// --- Siemens Structured Format ---
DATA_BLOCK "model_HS16_IW100"
{ S7_Optimized_Access := 'TRUE' }
VERSION : 0.1
NON_RETAIN
   VAR
      W_i : ARRAY[0..15, 0..39] OF REAL;
      W_f : ARRAY[0..15, 0..39] OF REAL;
      W_g : ARRAY[0..15, 0..39] OF REAL;
      W_o : ARRAY[0..15, 0..39] OF REAL;
      R_i : ARRAY[0..15, 0..15] OF REAL;
      R_f : ARRAY[0..15, 0..15] OF REAL;
      R_g : ARRAY[0..15, 0..15] OF REAL;
      R_o : ARRAY[0..15, 0..15] OF REAL;
      B_i : ARRAY[0..15] OF REAL;
      B_f : ARRAY[0..15] OF REAL;
      B_g : ARRAY[0..15] OF REAL;
      B_o : ARRAY[0..15] OF REAL;
      FC_W : ARRAY[0..39, 0..15] OF REAL;
      FC_B : ARRAY[0..39] OF REAL;
   END_VAR
BEGIN

      W_i[0,0] := 0.01364156;
      W_i[0,1] := 0.20536570;
      W_i[0,2] := -0.02245892;
      W_i[0,3] := 0.18291217;
      W_i[0,4] := 0.10548387;
      W_i[0,5] := 0.14748915;
      W_i[0,6] := 0.17824732;
      W_i[0,7] := 0.18831865;
      W_i[0,8] := 0.12917581;
      W_i[0,9] := -0.17035837;
      W_i[0,10] := 0.08922281;
      W_i[0,11] := -0.48598647;
      W_i[0,12] := -0.26934940;
      W_i[0,13] := -0.09021819;
      W_i[0,14] := 0.04866360;
      W_i[0,15] := 0.12027069;
      W_i[0,16] := 0.02211623;
      W_i[0,17] := -0.07331901;
      W_i[0,18] := 0.24969472;
      W_i[0,19] := 0.19951487;
      W_i[0,20] := -0.04635275;
      W_i[0,21] := -0.06017390;
      W_i[0,22] := 0.41972119;
      W_i[0,23] := -0.03179805;
      W_i[0,24] := 0.49648565;
      W_i[0,25] := 0.57860100;
      W_i[0,26] := -0.26113316;
      W_i[0,27] := -0.19300961;
      W_i[0,28] := 0.02716148;
      W_i[0,29] := -0.42831215;
      W_i[0,30] := 0.75518680;
      W_i[0,31] := -0.19160482;
      W_i[0,32] := 0.19652441;
      W_i[0,33] := 0.20859936;
      W_i[0,34] := 0.61514384;
      W_i[0,35] := -0.22654997;
      W_i[0,36] := -0.23919837;
      W_i[0,37] := -0.27295426;
      W_i[0,38] := 0.15717822;
      W_i[0,39] := 0.49166107;
      W_i[1,0] := -0.08388980;
      W_i[1,1] := 0.04137634;
      W_i[1,2] := 0.09732703;
      W_i[1,3] := -0.00114318;
      W_i[1,4] := 0.01266066;
      W_i[1,5] := 0.02146709;
      W_i[1,6] := 0.06203580;
      W_i[1,7] := -0.05510464;
      W_i[1,8] := 0.00995585;
      W_i[1,9] := -0.04009213;
      W_i[1,10] := -0.01534687;
      W_i[1,11] := -0.12621376;
      W_i[1,12] := -0.13568968;
      W_i[1,13] := -0.09674840;
      W_i[1,14] := -0.04467043;
      W_i[1,15] := -0.02089421;
      W_i[1,16] := -0.00725821;
      W_i[1,17] := 0.01724758;
      W_i[1,18] := 0.18129900;
      W_i[1,19] := 0.11187042;
      W_i[1,20] := 0.02454385;
      W_i[1,21] := -0.01102624;
      W_i[1,22] := 0.04567170;
      W_i[1,23] := -0.00008619;
      W_i[1,24] := -0.20038819;
      W_i[1,25] := -0.30851075;
      W_i[1,26] := 0.09543601;
      W_i[1,27] := -0.08277476;
      W_i[1,28] := 0.00373672;
      W_i[1,29] := -0.13582148;
      W_i[1,30] := 0.17890492;
      W_i[1,31] := 0.02590448;
      W_i[1,32] := 0.24079625;
      W_i[1,33] := -0.10525580;
      W_i[1,34] := -0.15286346;
      W_i[1,35] := -0.19629247;
      W_i[1,36] := -0.05740929;
      W_i[1,37] := 0.08565215;
      W_i[1,38] := 0.00725868;
      W_i[1,39] := 0.08298402;
      W_i[2,0] := -0.13536657;
      W_i[2,1] := 0.11532924;
      W_i[2,2] := 0.00179968;
      W_i[2,3] := -0.08932642;
      W_i[2,4] := 0.07508986;
      W_i[2,5] := -0.14212745;
      W_i[2,6] := -0.01394915;
      W_i[2,7] := -0.08767878;
      W_i[2,8] := 0.02846143;
      W_i[2,9] := 0.06891385;
      W_i[2,10] := 0.04481447;
      W_i[2,11] := -0.18693379;
      W_i[2,12] := 0.00844815;
      W_i[2,13] := -0.05949695;
      W_i[2,14] := 0.03289747;
      W_i[2,15] := 0.08402885;
      W_i[2,16] := 0.03656591;
      W_i[2,17] := 0.13008708;
      W_i[2,18] := -0.01728439;
      W_i[2,19] := -0.00760848;
      W_i[2,20] := -0.14490703;
      W_i[2,21] := 0.00184717;
      W_i[2,22] := -0.14345044;
      W_i[2,23] := -0.04114061;
      W_i[2,24] := 0.06368703;
      W_i[2,25] := -0.11341992;
      W_i[2,26] := -0.20044473;
      W_i[2,27] := -0.10808504;
      W_i[2,28] := -0.00091656;
      W_i[2,29] := -0.06285433;
      W_i[2,30] := 0.15420522;
      W_i[2,31] := -0.13147083;
      W_i[2,32] := -0.00983954;
      W_i[2,33] := -0.25118774;
      W_i[2,34] := -0.22324753;
      W_i[2,35] := -0.03245824;
      W_i[2,36] := 0.03434758;
      W_i[2,37] := -0.15230893;
      W_i[2,38] := 0.03214991;
      W_i[2,39] := 0.13666461;
      W_i[3,0] := -0.00015489;
      W_i[3,1] := -0.02602717;
      W_i[3,2] := 0.02940982;
      W_i[3,3] := 0.04201458;
      W_i[3,4] := 0.07303519;
      W_i[3,5] := 0.01782909;
      W_i[3,6] := -0.03795192;
      W_i[3,7] := -0.03116271;
      W_i[3,8] := 0.04315468;
      W_i[3,9] := -0.10355810;
      W_i[3,10] := 0.00910736;
      W_i[3,11] := 0.04493538;
      W_i[3,12] := 0.05511931;
      W_i[3,13] := 0.04794433;
      W_i[3,14] := -0.00690552;
      W_i[3,15] := 0.03096941;
      W_i[3,16] := 0.00754327;
      W_i[3,17] := 0.01626078;
      W_i[3,18] := -0.02028959;
      W_i[3,19] := -0.00735506;
      W_i[3,20] := -0.11980021;
      W_i[3,21] := -0.24100865;
      W_i[3,22] := 0.04234595;
      W_i[3,23] := -0.04032298;
      W_i[3,24] := -0.08977890;
      W_i[3,25] := 0.00863097;
      W_i[3,26] := -0.15812668;
      W_i[3,27] := 0.02937102;
      W_i[3,28] := 0.15920541;
      W_i[3,29] := -0.00798148;
      W_i[3,30] := -0.04935832;
      W_i[3,31] := -0.04004486;
      W_i[3,32] := -0.05156282;
      W_i[3,33] := -0.22839788;
      W_i[3,34] := 0.04730661;
      W_i[3,35] := -0.08628614;
      W_i[3,36] := 0.05156694;
      W_i[3,37] := 0.19403307;
      W_i[3,38] := 0.05496961;
      W_i[3,39] := -0.22899017;
      W_i[4,0] := -0.06762198;
      W_i[4,1] := 0.04105477;
      W_i[4,2] := 0.01412702;
      W_i[4,3] := -0.14503658;
      W_i[4,4] := 0.00052001;
      W_i[4,5] := -0.06361318;
      W_i[4,6] := 0.09927795;
      W_i[4,7] := 0.22318134;
      W_i[4,8] := 0.09787519;
      W_i[4,9] := 0.15435791;
      W_i[4,10] := -0.23381770;
      W_i[4,11] := -0.00151448;
      W_i[4,12] := -0.02443174;
      W_i[4,13] := -0.14362684;
      W_i[4,14] := 0.06250123;
      W_i[4,15] := -0.03108552;
      W_i[4,16] := -0.00760642;
      W_i[4,17] := -0.06110801;
      W_i[4,18] := 0.47297871;
      W_i[4,19] := 0.14145297;
      W_i[4,20] := -0.06666926;
      W_i[4,21] := 0.11880186;
      W_i[4,22] := 0.01305235;
      W_i[4,23] := -0.01088445;
      W_i[4,24] := 0.58226085;
      W_i[4,25] := 0.56463838;
      W_i[4,26] := -0.07272944;
      W_i[4,27] := -0.20381725;
      W_i[4,28] := 0.02941751;
      W_i[4,29] := 0.14696015;
      W_i[4,30] := -0.06698419;
      W_i[4,31] := -0.08342854;
      W_i[4,32] := 0.09379109;
      W_i[4,33] := 0.14583473;
      W_i[4,34] := -0.02093923;
      W_i[4,35] := -0.13240194;
      W_i[4,36] := -0.03764428;
      W_i[4,37] := -0.08758924;
      W_i[4,38] := -0.06055138;
      W_i[4,39] := 0.54854435;
      W_i[5,0] := -0.26418173;
      W_i[5,1] := 0.00919414;
      W_i[5,2] := 0.28921035;
      W_i[5,3] := 0.19848731;
      W_i[5,4] := 0.04857918;
      W_i[5,5] := -0.07696015;
      W_i[5,6] := -0.18773772;
      W_i[5,7] := -0.06413802;
      W_i[5,8] := -0.19999725;
      W_i[5,9] := 0.00090761;
      W_i[5,10] := 0.06217722;
      W_i[5,11] := 0.10535000;
      W_i[5,12] := -0.20478797;
      W_i[5,13] := 0.00378444;
      W_i[5,14] := -0.08047202;
      W_i[5,15] := 0.10188833;
      W_i[5,16] := -0.10373244;
      W_i[5,17] := 0.02060685;
      W_i[5,18] := 0.26179335;
      W_i[5,19] := -0.16465248;
      W_i[5,20] := -0.21371244;
      W_i[5,21] := 0.18068251;
      W_i[5,22] := -0.14789225;
      W_i[5,23] := -0.00876896;
      W_i[5,24] := 0.22973008;
      W_i[5,25] := 0.59550780;
      W_i[5,26] := 0.14612897;
      W_i[5,27] := -0.08599184;
      W_i[5,28] := -0.22050266;
      W_i[5,29] := -0.17621692;
      W_i[5,30] := -0.21464045;
      W_i[5,31] := -0.01781221;
      W_i[5,32] := -0.06129935;
      W_i[5,33] := 0.05988304;
      W_i[5,34] := 0.25511330;
      W_i[5,35] := -0.14653285;
      W_i[5,36] := -0.15237394;
      W_i[5,37] := -0.39873159;
      W_i[5,38] := 0.06444512;
      W_i[5,39] := -0.46595329;
      W_i[6,0] := -0.09987911;
      W_i[6,1] := -0.35666752;
      W_i[6,2] := -0.14997965;
      W_i[6,3] := -0.16122143;
      W_i[6,4] := -0.03222676;
      W_i[6,5] := -0.06696601;
      W_i[6,6] := -0.18053886;
      W_i[6,7] := -0.38125506;
      W_i[6,8] := 0.15195245;
      W_i[6,9] := -0.12253319;
      W_i[6,10] := -0.06935552;
      W_i[6,11] := -0.25237226;
      W_i[6,12] := -0.00955063;
      W_i[6,13] := -0.13364333;
      W_i[6,14] := 0.12441263;
      W_i[6,15] := -0.06698428;
      W_i[6,16] := 0.02953966;
      W_i[6,17] := -0.12817322;
      W_i[6,18] := 0.50510013;
      W_i[6,19] := -0.07000107;
      W_i[6,20] := 0.10518134;
      W_i[6,21] := -0.12933129;
      W_i[6,22] := 0.08060265;
      W_i[6,23] := 0.16216518;
      W_i[6,24] := 0.56379879;
      W_i[6,25] := 0.51589292;
      W_i[6,26] := -0.06017810;
      W_i[6,27] := 0.13627745;
      W_i[6,28] := 0.07406422;
      W_i[6,29] := -0.04566135;
      W_i[6,30] := 0.11365223;
      W_i[6,31] := -0.19966318;
      W_i[6,32] := 0.05134548;
      W_i[6,33] := -0.06383436;
      W_i[6,34] := 0.18601419;
      W_i[6,35] := -0.00495438;
      W_i[6,36] := -0.01991113;
      W_i[6,37] := 0.13569827;
      W_i[6,38] := 0.10721204;
      W_i[6,39] := -0.19543035;
      W_i[7,0] := 0.11805627;
      W_i[7,1] := 0.06404518;
      W_i[7,2] := 0.26091906;
      W_i[7,3] := -0.13242221;
      W_i[7,4] := 0.04345745;
      W_i[7,5] := 0.06463753;
      W_i[7,6] := 0.14174174;
      W_i[7,7] := 0.17861204;
      W_i[7,8] := 0.14897110;
      W_i[7,9] := -0.10119636;
      W_i[7,10] := -0.21339175;
      W_i[7,11] := -0.29427007;
      W_i[7,12] := -0.12524955;
      W_i[7,13] := -0.22747980;
      W_i[7,14] := -0.08303443;
      W_i[7,15] := 0.15086012;
      W_i[7,16] := -0.02865510;
      W_i[7,17] := 0.14286377;
      W_i[7,18] := 0.06569705;
      W_i[7,19] := 0.17024888;
      W_i[7,20] := 0.16341139;
      W_i[7,21] := -0.08116058;
      W_i[7,22] := 0.28119785;
      W_i[7,23] := -0.24578308;
      W_i[7,24] := 0.46118793;
      W_i[7,25] := 0.87448853;
      W_i[7,26] := -0.21451366;
      W_i[7,27] := -0.03196089;
      W_i[7,28] := 0.11030190;
      W_i[7,29] := 0.08675592;
      W_i[7,30] := 0.63182199;
      W_i[7,31] := 0.09978309;
      W_i[7,32] := -0.11112560;
      W_i[7,33] := 0.14244974;
      W_i[7,34] := 0.87706214;
      W_i[7,35] := 0.04549777;
      W_i[7,36] := 0.01875403;
      W_i[7,37] := 0.19351047;
      W_i[7,38] := 0.04132079;
      W_i[7,39] := 0.30163178;
      W_i[8,0] := 0.00448507;
      W_i[8,1] := 0.00593045;
      W_i[8,2] := 0.05385492;
      W_i[8,3] := 0.23692533;
      W_i[8,4] := 0.13600577;
      W_i[8,5] := -0.13479330;
      W_i[8,6] := 0.05155064;
      W_i[8,7] := -0.18396251;
      W_i[8,8] := -0.04175631;
      W_i[8,9] := 0.02508196;
      W_i[8,10] := 0.08028799;
      W_i[8,11] := -0.09709663;
      W_i[8,12] := -0.24632221;
      W_i[8,13] := -0.09933189;
      W_i[8,14] := -0.13090380;
      W_i[8,15] := 0.08873132;
      W_i[8,16] := -0.15212885;
      W_i[8,17] := 0.09358153;
      W_i[8,18] := -0.04925272;
      W_i[8,19] := -0.20840898;
      W_i[8,20] := -0.08381097;
      W_i[8,21] := 0.06258945;
      W_i[8,22] := -0.07553499;
      W_i[8,23] := -0.05963936;
      W_i[8,24] := 0.35542277;
      W_i[8,25] := 0.42086950;
      W_i[8,26] := 0.08319889;
      W_i[8,27] := -0.18197235;
      W_i[8,28] := 0.06505518;
      W_i[8,29] := 0.07391432;
      W_i[8,30] := 0.12715283;
      W_i[8,31] := -0.13722460;
      W_i[8,32] := 0.24457708;
      W_i[8,33] := 0.17096752;
      W_i[8,34] := -0.13092747;
      W_i[8,35] := 0.11238978;
      W_i[8,36] := -0.01007767;
      W_i[8,37] := 0.04878357;
      W_i[8,38] := -0.09178042;
      W_i[8,39] := 0.70590818;
      W_i[9,0] := 0.13898331;
      W_i[9,1] := 0.21558045;
      W_i[9,2] := -0.01587300;
      W_i[9,3] := -0.02008759;
      W_i[9,4] := 0.14031912;
      W_i[9,5] := 0.14432517;
      W_i[9,6] := 0.22022982;
      W_i[9,7] := 0.11039817;
      W_i[9,8] := -0.01799948;
      W_i[9,9] := 0.01688460;
      W_i[9,10] := 0.08939565;
      W_i[9,11] := 0.15729012;
      W_i[9,12] := -0.16055229;
      W_i[9,13] := 0.07329134;
      W_i[9,14] := 0.03671210;
      W_i[9,15] := 0.07092312;
      W_i[9,16] := -0.01012265;
      W_i[9,17] := 0.03808835;
      W_i[9,18] := -0.00362916;
      W_i[9,19] := -0.00791038;
      W_i[9,20] := 0.13901256;
      W_i[9,21] := -0.05212758;
      W_i[9,22] := -0.13945961;
      W_i[9,23] := 0.01820100;
      W_i[9,24] := -0.28223145;
      W_i[9,25] := -0.05683075;
      W_i[9,26] := -0.06647032;
      W_i[9,27] := 0.11427623;
      W_i[9,28] := -0.05756322;
      W_i[9,29] := 0.25496486;
      W_i[9,30] := -0.41661564;
      W_i[9,31] := 0.03821095;
      W_i[9,32] := -0.24074574;
      W_i[9,33] := -0.01633074;
      W_i[9,34] := -0.30772033;
      W_i[9,35] := -0.30636224;
      W_i[9,36] := -0.00646075;
      W_i[9,37] := -0.10956979;
      W_i[9,38] := 0.04284515;
      W_i[9,39] := 0.06388737;
      W_i[10,0] := 0.15491682;
      W_i[10,1] := 0.06016659;
      W_i[10,2] := 0.08790326;
      W_i[10,3] := 0.04701571;
      W_i[10,4] := -0.21938066;
      W_i[10,5] := -0.00418864;
      W_i[10,6] := -0.14329411;
      W_i[10,7] := -0.13763005;
      W_i[10,8] := -0.07890343;
      W_i[10,9] := 0.10256134;
      W_i[10,10] := -0.02710062;
      W_i[10,11] := -0.20991582;
      W_i[10,12] := 0.43801337;
      W_i[10,13] := 0.07667056;
      W_i[10,14] := -0.05265489;
      W_i[10,15] := 0.09571737;
      W_i[10,16] := -0.14256968;
      W_i[10,17] := 0.00645238;
      W_i[10,18] := 0.08263779;
      W_i[10,19] := -0.13588426;
      W_i[10,20] := 0.17050405;
      W_i[10,21] := 0.34270245;
      W_i[10,22] := 0.12177468;
      W_i[10,23] := 0.03954393;
      W_i[10,24] := 0.78272396;
      W_i[10,25] := 0.62249583;
      W_i[10,26] := -0.04197677;
      W_i[10,27] := -0.01324140;
      W_i[10,28] := -0.11742962;
      W_i[10,29] := 0.03315270;
      W_i[10,30] := 0.43726227;
      W_i[10,31] := -0.01188345;
      W_i[10,32] := 0.02015782;
      W_i[10,33] := 0.26254645;
      W_i[10,34] := 0.31372723;
      W_i[10,35] := 0.13515088;
      W_i[10,36] := -0.13856903;
      W_i[10,37] := -0.07906500;
      W_i[10,38] := 0.04151168;
      W_i[10,39] := 0.58438212;
      W_i[11,0] := -0.03692184;
      W_i[11,1] := 0.08602915;
      W_i[11,2] := 0.04734402;
      W_i[11,3] := 0.15488507;
      W_i[11,4] := 0.02953814;
      W_i[11,5] := -0.03516553;
      W_i[11,6] := -0.03630468;
      W_i[11,7] := 0.22055247;
      W_i[11,8] := 0.05422686;
      W_i[11,9] := -0.19223477;
      W_i[11,10] := 0.15922990;
      W_i[11,11] := -0.50660896;
      W_i[11,12] := 0.21863456;
      W_i[11,13] := 0.06115106;
      W_i[11,14] := 0.05269584;
      W_i[11,15] := 0.01791226;
      W_i[11,16] := -0.08076685;
      W_i[11,17] := -0.00192191;
      W_i[11,18] := 0.20004040;
      W_i[11,19] := -0.02625836;
      W_i[11,20] := 0.02325124;
      W_i[11,21] := 0.02411360;
      W_i[11,22] := -0.03470324;
      W_i[11,23] := 0.02441446;
      W_i[11,24] := 0.01363192;
      W_i[11,25] := -0.20787865;
      W_i[11,26] := -0.09482310;
      W_i[11,27] := 0.05317536;
      W_i[11,28] := 0.01368785;
      W_i[11,29] := 0.24679546;
      W_i[11,30] := 0.09310606;
      W_i[11,31] := 0.02022941;
      W_i[11,32] := 0.25092661;
      W_i[11,33] := -0.02307699;
      W_i[11,34] := -0.18370298;
      W_i[11,35] := 0.24884717;
      W_i[11,36] := -0.08544295;
      W_i[11,37] := -0.04159483;
      W_i[11,38] := 0.12627473;
      W_i[11,39] := 0.57147032;
      W_i[12,0] := 0.26667652;
      W_i[12,1] := 0.18141651;
      W_i[12,2] := -0.04977122;
      W_i[12,3] := 0.09079568;
      W_i[12,4] := 0.22469823;
      W_i[12,5] := -0.13473749;
      W_i[12,6] := 0.22730011;
      W_i[12,7] := -0.10648373;
      W_i[12,8] := 0.00375756;
      W_i[12,9] := 0.14409521;
      W_i[12,10] := -0.04439257;
      W_i[12,11] := 0.01341529;
      W_i[12,12] := 0.05264389;
      W_i[12,13] := 0.14714998;
      W_i[12,14] := 0.02812583;
      W_i[12,15] := 0.09371702;
      W_i[12,16] := -0.01640923;
      W_i[12,17] := -0.00820156;
      W_i[12,18] := -0.02099935;
      W_i[12,19] := 0.03455377;
      W_i[12,20] := -0.00376845;
      W_i[12,21] := 0.01287318;
      W_i[12,22] := 0.27967688;
      W_i[12,23] := 0.32648781;
      W_i[12,24] := -0.04639676;
      W_i[12,25] := -0.12604533;
      W_i[12,26] := -0.05218698;
      W_i[12,27] := 0.19303280;
      W_i[12,28] := -0.02861599;
      W_i[12,29] := 0.07526918;
      W_i[12,30] := 0.27195212;
      W_i[12,31] := -0.24740550;
      W_i[12,32] := 0.12962508;
      W_i[12,33] := -0.02061021;
      W_i[12,34] := -0.38526946;
      W_i[12,35] := -0.44955108;
      W_i[12,36] := 0.17704585;
      W_i[12,37] := -0.58847874;
      W_i[12,38] := 0.02093910;
      W_i[12,39] := -0.07715891;
      W_i[13,0] := 0.02638375;
      W_i[13,1] := 0.04267908;
      W_i[13,2] := -0.04100905;
      W_i[13,3] := 0.02433234;
      W_i[13,4] := 0.19633174;
      W_i[13,5] := 0.09253235;
      W_i[13,6] := 0.18767522;
      W_i[13,7] := -0.09313158;
      W_i[13,8] := 0.06435700;
      W_i[13,9] := -0.02719559;
      W_i[13,10] := 0.11561871;
      W_i[13,11] := -0.12066963;
      W_i[13,12] := -0.27772844;
      W_i[13,13] := -0.00763909;
      W_i[13,14] := 0.07759997;
      W_i[13,15] := 0.01202866;
      W_i[13,16] := 0.07374192;
      W_i[13,17] := 0.03084671;
      W_i[13,18] := -0.03566260;
      W_i[13,19] := 0.21000803;
      W_i[13,20] := -0.08411094;
      W_i[13,21] := -0.21406713;
      W_i[13,22] := 0.03648549;
      W_i[13,23] := -0.03847607;
      W_i[13,24] := 0.70946354;
      W_i[13,25] := 0.49792659;
      W_i[13,26] := -0.08645725;
      W_i[13,27] := 0.15172665;
      W_i[13,28] := -0.01545484;
      W_i[13,29] := 0.07564367;
      W_i[13,30] := 0.04488704;
      W_i[13,31] := -0.05433368;
      W_i[13,32] := -0.12254967;
      W_i[13,33] := 0.05323875;
      W_i[13,34] := 0.28031611;
      W_i[13,35] := -0.31686431;
      W_i[13,36] := 0.08479394;
      W_i[13,37] := -0.18495709;
      W_i[13,38] := 0.10758790;
      W_i[13,39] := 0.68741995;
      W_i[14,0] := -0.17416088;
      W_i[14,1] := 0.01005446;
      W_i[14,2] := -0.26855752;
      W_i[14,3] := -0.62796623;
      W_i[14,4] := 0.06820592;
      W_i[14,5] := -0.16153112;
      W_i[14,6] := 0.04283209;
      W_i[14,7] := -0.29056939;
      W_i[14,8] := -0.67249602;
      W_i[14,9] := -0.34167016;
      W_i[14,10] := 0.09426845;
      W_i[14,11] := -0.10104106;
      W_i[14,12] := 0.10796092;
      W_i[14,13] := -0.18351264;
      W_i[14,14] := 0.00065603;
      W_i[14,15] := -0.06139126;
      W_i[14,16] := -0.11547680;
      W_i[14,17] := 0.04488576;
      W_i[14,18] := -0.15664500;
      W_i[14,19] := 0.00779267;
      W_i[14,20] := -0.01367023;
      W_i[14,21] := -0.02746255;
      W_i[14,22] := -0.06486769;
      W_i[14,23] := 0.17152609;
      W_i[14,24] := -0.10990940;
      W_i[14,25] := -0.08006914;
      W_i[14,26] := -0.25285053;
      W_i[14,27] := 0.06160279;
      W_i[14,28] := 0.17719766;
      W_i[14,29] := 0.14922956;
      W_i[14,30] := 0.00092594;
      W_i[14,31] := -0.11380912;
      W_i[14,32] := -0.09275766;
      W_i[14,33] := -0.05691696;
      W_i[14,34] := -0.20431529;
      W_i[14,35] := -0.06423868;
      W_i[14,36] := -0.08797362;
      W_i[14,37] := -0.07569788;
      W_i[14,38] := 0.23112053;
      W_i[14,39] := 0.00680392;
      W_i[15,0] := 0.02184013;
      W_i[15,1] := 0.18801539;
      W_i[15,2] := 0.06529985;
      W_i[15,3] := -0.13560045;
      W_i[15,4] := 0.14931200;
      W_i[15,5] := -0.07038850;
      W_i[15,6] := -0.03877895;
      W_i[15,7] := 0.08169580;
      W_i[15,8] := 0.04022081;
      W_i[15,9] := 0.16485462;
      W_i[15,10] := 0.02359114;
      W_i[15,11] := -0.06464480;
      W_i[15,12] := -0.13054129;
      W_i[15,13] := 0.14513132;
      W_i[15,14] := -0.00291753;
      W_i[15,15] := 0.00511506;
      W_i[15,16] := 0.04386861;
      W_i[15,17] := -0.14875175;
      W_i[15,18] := -0.02457544;
      W_i[15,19] := 0.07704978;
      W_i[15,20] := -0.04825005;
      W_i[15,21] := 0.03190987;
      W_i[15,22] := -0.09410153;
      W_i[15,23] := -0.16679235;
      W_i[15,24] := -0.46764547;
      W_i[15,25] := -0.44318548;
      W_i[15,26] := -0.05940514;
      W_i[15,27] := 0.05163483;
      W_i[15,28] := -0.03008339;
      W_i[15,29] := 0.21256405;
      W_i[15,30] := -0.05510921;
      W_i[15,31] := -0.09820909;
      W_i[15,32] := 0.21482152;
      W_i[15,33] := 0.30279014;
      W_i[15,34] := -0.06246981;
      W_i[15,35] := 0.01027228;
      W_i[15,36] := -0.09376621;
      W_i[15,37] := -0.02936010;
      W_i[15,38] := -0.47935137;
      W_i[15,39] := 0.05519279;
      W_f[0,0] := 0.05364275;
      W_f[0,1] := 0.09687193;
      W_f[0,2] := -0.03420604;
      W_f[0,3] := 0.09112332;
      W_f[0,4] := 0.01952212;
      W_f[0,5] := -0.00599490;
      W_f[0,6] := -0.02583287;
      W_f[0,7] := 0.01641575;
      W_f[0,8] := 0.00249371;
      W_f[0,9] := -0.03082566;
      W_f[0,10] := 0.03822958;
      W_f[0,11] := -0.20525688;
      W_f[0,12] := 0.15610816;
      W_f[0,13] := 0.01319965;
      W_f[0,14] := -0.00955972;
      W_f[0,15] := -0.01736578;
      W_f[0,16] := -0.01232213;
      W_f[0,17] := -0.07847971;
      W_f[0,18] := 0.03267125;
      W_f[0,19] := 0.02281226;
      W_f[0,20] := -0.00946235;
      W_f[0,21] := -0.04914912;
      W_f[0,22] := -0.05509606;
      W_f[0,23] := -0.04103199;
      W_f[0,24] := 0.49705139;
      W_f[0,25] := 0.41528228;
      W_f[0,26] := -0.10808732;
      W_f[0,27] := -0.04818393;
      W_f[0,28] := 0.06444012;
      W_f[0,29] := -0.15780614;
      W_f[0,30] := 0.10075731;
      W_f[0,31] := -0.03347747;
      W_f[0,32] := 0.13920051;
      W_f[0,33] := -0.07730422;
      W_f[0,34] := 0.22286199;
      W_f[0,35] := 0.09730371;
      W_f[0,36] := 0.01644731;
      W_f[0,37] := -0.14617991;
      W_f[0,38] := -0.03747354;
      W_f[0,39] := 0.08508820;
      W_f[1,0] := -0.03535822;
      W_f[1,1] := -0.47124356;
      W_f[1,2] := -0.14644240;
      W_f[1,3] := 0.07842869;
      W_f[1,4] := -0.00283514;
      W_f[1,5] := 0.13242532;
      W_f[1,6] := -0.17787769;
      W_f[1,7] := 0.03437876;
      W_f[1,8] := -0.30326170;
      W_f[1,9] := 0.03390699;
      W_f[1,10] := 0.04835700;
      W_f[1,11] := 0.39755464;
      W_f[1,12] := 0.22270909;
      W_f[1,13] := 0.21808504;
      W_f[1,14] := -0.11776564;
      W_f[1,15] := 0.10067453;
      W_f[1,16] := -0.36373556;
      W_f[1,17] := 0.18559641;
      W_f[1,18] := 0.40969753;
      W_f[1,19] := 0.12707092;
      W_f[1,20] := 0.29767519;
      W_f[1,21] := -0.16713570;
      W_f[1,22] := -0.17408817;
      W_f[1,23] := 0.12793775;
      W_f[1,24] := -0.53485709;
      W_f[1,25] := -0.56272870;
      W_f[1,26] := 0.05998780;
      W_f[1,27] := 0.01051460;
      W_f[1,28] := -0.12135706;
      W_f[1,29] := 0.13744721;
      W_f[1,30] := -0.09007506;
      W_f[1,31] := -0.00778998;
      W_f[1,32] := 0.11112776;
      W_f[1,33] := -0.16928056;
      W_f[1,34] := 0.31107175;
      W_f[1,35] := 0.19411123;
      W_f[1,36] := -0.06959353;
      W_f[1,37] := -0.25251710;
      W_f[1,38] := 0.34865397;
      W_f[1,39] := 0.05812330;
      W_f[2,0] := -0.03221922;
      W_f[2,1] := 0.12347551;
      W_f[2,2] := -0.06227477;
      W_f[2,3] := 0.20185524;
      W_f[2,4] := 0.00543583;
      W_f[2,5] := 0.03781491;
      W_f[2,6] := -0.00314693;
      W_f[2,7] := 0.04292703;
      W_f[2,8] := -0.00575330;
      W_f[2,9] := -0.08594991;
      W_f[2,10] := -0.01364730;
      W_f[2,11] := -0.17743753;
      W_f[2,12] := -0.00461064;
      W_f[2,13] := -0.05826429;
      W_f[2,14] := 0.06936967;
      W_f[2,15] := 0.02028695;
      W_f[2,16] := 0.00601915;
      W_f[2,17] := 0.02327365;
      W_f[2,18] := -0.03857812;
      W_f[2,19] := -0.08794222;
      W_f[2,20] := 0.01833609;
      W_f[2,21] := 0.03344638;
      W_f[2,22] := -0.09674103;
      W_f[2,23] := 0.03481310;
      W_f[2,24] := -0.20710675;
      W_f[2,25] := -0.12916997;
      W_f[2,26] := 0.00745270;
      W_f[2,27] := -0.01033618;
      W_f[2,28] := 0.07703895;
      W_f[2,29] := 0.08949607;
      W_f[2,30] := -0.07744866;
      W_f[2,31] := -0.00363669;
      W_f[2,32] := -0.10897757;
      W_f[2,33] := 0.05933027;
      W_f[2,34] := 0.12423457;
      W_f[2,35] := -0.08927383;
      W_f[2,36] := -0.00645528;
      W_f[2,37] := 0.19684052;
      W_f[2,38] := -0.12688994;
      W_f[2,39] := 0.15507455;
      W_f[3,0] := -0.15219240;
      W_f[3,1] := -0.09112048;
      W_f[3,2] := -0.13655797;
      W_f[3,3] := 0.09398650;
      W_f[3,4] := -0.38095236;
      W_f[3,5] := 0.07147726;
      W_f[3,6] := 0.27381626;
      W_f[3,7] := -0.03780884;
      W_f[3,8] := -0.09247751;
      W_f[3,9] := 0.32965410;
      W_f[3,10] := -0.21033977;
      W_f[3,11] := -0.01770502;
      W_f[3,12] := -0.16563010;
      W_f[3,13] := -0.09659225;
      W_f[3,14] := -0.14708968;
      W_f[3,15] := -0.04307340;
      W_f[3,16] := -0.04020571;
      W_f[3,17] := -0.15388337;
      W_f[3,18] := 0.04561477;
      W_f[3,19] := -0.03800451;
      W_f[3,20] := -0.11640513;
      W_f[3,21] := 0.10628393;
      W_f[3,22] := 0.13051899;
      W_f[3,23] := 0.15934397;
      W_f[3,24] := -0.49496132;
      W_f[3,25] := -0.46555015;
      W_f[3,26] := 0.07467606;
      W_f[3,27] := 0.05813665;
      W_f[3,28] := -0.45595208;
      W_f[3,29] := 0.13731937;
      W_f[3,30] := -0.04639205;
      W_f[3,31] := 0.20856442;
      W_f[3,32] := 0.23197061;
      W_f[3,33] := -0.09503688;
      W_f[3,34] := 0.22798222;
      W_f[3,35] := -0.10183924;
      W_f[3,36] := 0.24291022;
      W_f[3,37] := 0.09243517;
      W_f[3,38] := -0.01472234;
      W_f[3,39] := 0.84467447;
      W_f[4,0] := 0.02846950;
      W_f[4,1] := 0.06578626;
      W_f[4,2] := 0.00272045;
      W_f[4,3] := 0.02383544;
      W_f[4,4] := -0.04941020;
      W_f[4,5] := 0.03107557;
      W_f[4,6] := 0.04498140;
      W_f[4,7] := 0.00715393;
      W_f[4,8] := -0.00156786;
      W_f[4,9] := 0.01842991;
      W_f[4,10] := -0.02190995;
      W_f[4,11] := 0.00170467;
      W_f[4,12] := -0.11754189;
      W_f[4,13] := -0.00572082;
      W_f[4,14] := -0.02148229;
      W_f[4,15] := -0.02594547;
      W_f[4,16] := -0.06025682;
      W_f[4,17] := -0.08476730;
      W_f[4,18] := 0.07604560;
      W_f[4,19] := 0.05858169;
      W_f[4,20] := 0.05974808;
      W_f[4,21] := 0.24128842;
      W_f[4,22] := 0.16804713;
      W_f[4,23] := -0.03820573;
      W_f[4,24] := 0.48765618;
      W_f[4,25] := 0.57080442;
      W_f[4,26] := -0.00810769;
      W_f[4,27] := -0.18718927;
      W_f[4,28] := 0.06110260;
      W_f[4,29] := -0.09344726;
      W_f[4,30] := 0.46467450;
      W_f[4,31] := 0.05612971;
      W_f[4,32] := 0.03677486;
      W_f[4,33] := 0.11877728;
      W_f[4,34] := 0.03321171;
      W_f[4,35] := 0.29353175;
      W_f[4,36] := 0.05504971;
      W_f[4,37] := 0.10279266;
      W_f[4,38] := -0.00283241;
      W_f[4,39] := 0.06622307;
      W_f[5,0] := 0.11376505;
      W_f[5,1] := 0.04806940;
      W_f[5,2] := -0.10279931;
      W_f[5,3] := -0.16593064;
      W_f[5,4] := 0.00000844;
      W_f[5,5] := 0.02789909;
      W_f[5,6] := 0.04521109;
      W_f[5,7] := 0.02275284;
      W_f[5,8] := -0.02738458;
      W_f[5,9] := 0.06878603;
      W_f[5,10] := -0.01160701;
      W_f[5,11] := -0.05195494;
      W_f[5,12] := -0.10548418;
      W_f[5,13] := 0.01500680;
      W_f[5,14] := 0.08265527;
      W_f[5,15] := 0.00386744;
      W_f[5,16] := 0.05198263;
      W_f[5,17] := 0.02937749;
      W_f[5,18] := 0.06512810;
      W_f[5,19] := 0.03703250;
      W_f[5,20] := 0.06421617;
      W_f[5,21] := -0.01455062;
      W_f[5,22] := 0.19789651;
      W_f[5,23] := -0.03008014;
      W_f[5,24] := 0.34697571;
      W_f[5,25] := 0.65106732;
      W_f[5,26] := -0.00135605;
      W_f[5,27] := 0.05647351;
      W_f[5,28] := 0.09934321;
      W_f[5,29] := -0.13159826;
      W_f[5,30] := 0.01969404;
      W_f[5,31] := 0.03655320;
      W_f[5,32] := -0.05406484;
      W_f[5,33] := -0.11042146;
      W_f[5,34] := 0.09479982;
      W_f[5,35] := 0.04922118;
      W_f[5,36] := 0.04102103;
      W_f[5,37] := 0.20328595;
      W_f[5,38] := 0.09994788;
      W_f[5,39] := 0.16133195;
      W_f[6,0] := -0.03485869;
      W_f[6,1] := -0.00908120;
      W_f[6,2] := -0.03699812;
      W_f[6,3] := -0.03682025;
      W_f[6,4] := 0.09187597;
      W_f[6,5] := 0.05246547;
      W_f[6,6] := 0.12492345;
      W_f[6,7] := -0.00999346;
      W_f[6,8] := -0.08344354;
      W_f[6,9] := 0.07932125;
      W_f[6,10] := 0.03438351;
      W_f[6,11] := -0.06988891;
      W_f[6,12] := 0.03135443;
      W_f[6,13] := 0.00137540;
      W_f[6,14] := 0.03249843;
      W_f[6,15] := -0.01266906;
      W_f[6,16] := -0.00345383;
      W_f[6,17] := -0.07384243;
      W_f[6,18] := -0.04767740;
      W_f[6,19] := 0.00589593;
      W_f[6,20] := 0.04428503;
      W_f[6,21] := 0.05965255;
      W_f[6,22] := 0.13275859;
      W_f[6,23] := -0.07216866;
      W_f[6,24] := 0.32743850;
      W_f[6,25] := 0.41480702;
      W_f[6,26] := 0.00211261;
      W_f[6,27] := -0.02340442;
      W_f[6,28] := -0.04405304;
      W_f[6,29] := 0.02433619;
      W_f[6,30] := -0.18997696;
      W_f[6,31] := 0.13028599;
      W_f[6,32] := 0.16898793;
      W_f[6,33] := 0.09330611;
      W_f[6,34] := 0.04484965;
      W_f[6,35] := -0.08660950;
      W_f[6,36] := -0.02266579;
      W_f[6,37] := 0.11412326;
      W_f[6,38] := 0.07686570;
      W_f[6,39] := -0.11869525;
      W_f[7,0] := -0.00221147;
      W_f[7,1] := 0.10511280;
      W_f[7,2] := -0.07019065;
      W_f[7,3] := -0.01243510;
      W_f[7,4] := 0.02943816;
      W_f[7,5] := 0.06614972;
      W_f[7,6] := 0.04611924;
      W_f[7,7] := 0.02763495;
      W_f[7,8] := -0.01057697;
      W_f[7,9] := -0.02540869;
      W_f[7,10] := -0.00237630;
      W_f[7,11] := -0.14796597;
      W_f[7,12] := 0.04395492;
      W_f[7,13] := 0.07364006;
      W_f[7,14] := -0.03409544;
      W_f[7,15] := -0.07690118;
      W_f[7,16] := 0.00728678;
      W_f[7,17] := 0.07319640;
      W_f[7,18] := 0.06380690;
      W_f[7,19] := 0.00555583;
      W_f[7,20] := -0.01266172;
      W_f[7,21] := 0.05246431;
      W_f[7,22] := 0.13432735;
      W_f[7,23] := 0.00786275;
      W_f[7,24] := 0.36037040;
      W_f[7,25] := 0.63975710;
      W_f[7,26] := -0.14318357;
      W_f[7,27] := 0.02217500;
      W_f[7,28] := 0.03329759;
      W_f[7,29] := 0.02024308;
      W_f[7,30] := 0.06194379;
      W_f[7,31] := -0.03574094;
      W_f[7,32] := 0.27383688;
      W_f[7,33] := 0.09022309;
      W_f[7,34] := 0.72298384;
      W_f[7,35] := -0.13958853;
      W_f[7,36] := -0.05832926;
      W_f[7,37] := 0.05806842;
      W_f[7,38] := 0.01794156;
      W_f[7,39] := 0.00930902;
      W_f[8,0] := -0.00069194;
      W_f[8,1] := 0.09570718;
      W_f[8,2] := -0.13032150;
      W_f[8,3] := -0.00169487;
      W_f[8,4] := 0.05343744;
      W_f[8,5] := 0.05416366;
      W_f[8,6] := 0.00489102;
      W_f[8,7] := 0.04302023;
      W_f[8,8] := 0.02923981;
      W_f[8,9] := -0.03308041;
      W_f[8,10] := 0.02764279;
      W_f[8,11] := -0.08082840;
      W_f[8,12] := -0.04773318;
      W_f[8,13] := -0.02026195;
      W_f[8,14] := -0.02248771;
      W_f[8,15] := -0.14968230;
      W_f[8,16] := 0.10387620;
      W_f[8,17] := 0.02660801;
      W_f[8,18] := 0.02133987;
      W_f[8,19] := 0.06662087;
      W_f[8,20] := 0.02782230;
      W_f[8,21] := 0.01667393;
      W_f[8,22] := 0.29885378;
      W_f[8,23] := -0.04644651;
      W_f[8,24] := 0.36805248;
      W_f[8,25] := 0.58228642;
      W_f[8,26] := -0.01743001;
      W_f[8,27] := -0.01691605;
      W_f[8,28] := 0.01118935;
      W_f[8,29] := -0.00426544;
      W_f[8,30] := 0.17033555;
      W_f[8,31] := -0.03053380;
      W_f[8,32] := 0.12107975;
      W_f[8,33] := -0.06191333;
      W_f[8,34] := 0.74060959;
      W_f[8,35] := -0.07475549;
      W_f[8,36] := -0.02023359;
      W_f[8,37] := 0.02331678;
      W_f[8,38] := -0.03007067;
      W_f[8,39] := -0.05748938;
      W_f[9,0] := -0.10508082;
      W_f[9,1] := -0.04133019;
      W_f[9,2] := -0.06146885;
      W_f[9,3] := 0.03741426;
      W_f[9,4] := -0.08707085;
      W_f[9,5] := -0.06223321;
      W_f[9,6] := -0.18814664;
      W_f[9,7] := -0.11111913;
      W_f[9,8] := -0.13546698;
      W_f[9,9] := -0.00564482;
      W_f[9,10] := -0.01552745;
      W_f[9,11] := -0.17684816;
      W_f[9,12] := 0.03565479;
      W_f[9,13] := -0.08725277;
      W_f[9,14] := -0.00522599;
      W_f[9,15] := -0.10947887;
      W_f[9,16] := 0.01476094;
      W_f[9,17] := -0.05979283;
      W_f[9,18] := -0.00063397;
      W_f[9,19] := 0.06166672;
      W_f[9,20] := -0.10422222;
      W_f[9,21] := 0.00166027;
      W_f[9,22] := -0.27992189;
      W_f[9,23] := -0.03734995;
      W_f[9,24] := 0.12155679;
      W_f[9,25] := -0.06815521;
      W_f[9,26] := -0.01121978;
      W_f[9,27] := -0.01608659;
      W_f[9,28] := 0.04067907;
      W_f[9,29] := -0.06756267;
      W_f[9,30] := 0.05508788;
      W_f[9,31] := -0.09057643;
      W_f[9,32] := -0.07261790;
      W_f[9,33] := -0.13291492;
      W_f[9,34] := -0.02277668;
      W_f[9,35] := 0.19900511;
      W_f[9,36] := -0.00467835;
      W_f[9,37] := -0.18864036;
      W_f[9,38] := 0.01334353;
      W_f[9,39] := -0.01253361;
      W_f[10,0] := -0.00524171;
      W_f[10,1] := 0.10620133;
      W_f[10,2] := -0.06919775;
      W_f[10,3] := -0.00134773;
      W_f[10,4] := -0.01228707;
      W_f[10,5] := 0.01736076;
      W_f[10,6] := 0.03687445;
      W_f[10,7] := 0.02915340;
      W_f[10,8] := 0.06300525;
      W_f[10,9] := -0.06548626;
      W_f[10,10] := 0.05580841;
      W_f[10,11] := -0.10701931;
      W_f[10,12] := -0.02223501;
      W_f[10,13] := 0.00853262;
      W_f[10,14] := 0.03023283;
      W_f[10,15] := -0.06348655;
      W_f[10,16] := 0.04187576;
      W_f[10,17] := 0.00731900;
      W_f[10,18] := 0.08542238;
      W_f[10,19] := 0.00890474;
      W_f[10,20] := 0.07895420;
      W_f[10,21] := 0.07658880;
      W_f[10,22] := 0.32859516;
      W_f[10,23] := -0.03547200;
      W_f[10,24] := 0.30065846;
      W_f[10,25] := 0.61635405;
      W_f[10,26] := 0.05265321;
      W_f[10,27] := 0.01765742;
      W_f[10,28] := 0.11246407;
      W_f[10,29] := 0.15208840;
      W_f[10,30] := 0.36211643;
      W_f[10,31] := -0.00268147;
      W_f[10,32] := 0.04235294;
      W_f[10,33] := 0.04691185;
      W_f[10,34] := 0.35568959;
      W_f[10,35] := 0.18353109;
      W_f[10,36] := 0.01559761;
      W_f[10,37] := 0.06422969;
      W_f[10,38] := -0.05459329;
      W_f[10,39] := 0.00331264;
      W_f[11,0] := 0.05995931;
      W_f[11,1] := -0.09904456;
      W_f[11,2] := -0.08644266;
      W_f[11,3] := -0.15029024;
      W_f[11,4] := 0.04589326;
      W_f[11,5] := 0.01600008;
      W_f[11,6] := 0.03320405;
      W_f[11,7] := 0.13276693;
      W_f[11,8] := 0.02298770;
      W_f[11,9] := -0.13637532;
      W_f[11,10] := -0.05902323;
      W_f[11,11] := 0.18438902;
      W_f[11,12] := 0.02477853;
      W_f[11,13] := 0.01040439;
      W_f[11,14] := -0.07367453;
      W_f[11,15] := 0.00079368;
      W_f[11,16] := 0.03881615;
      W_f[11,17] := 0.07118577;
      W_f[11,18] := -0.02313377;
      W_f[11,19] := 0.18068580;
      W_f[11,20] := -0.04932791;
      W_f[11,21] := 0.06971975;
      W_f[11,22] := -0.34139532;
      W_f[11,23] := 0.05619354;
      W_f[11,24] := -0.39076003;
      W_f[11,25] := -0.13438395;
      W_f[11,26] := 0.07639978;
      W_f[11,27] := 0.02963847;
      W_f[11,28] := 0.00480400;
      W_f[11,29] := 0.41879687;
      W_f[11,30] := -0.23149464;
      W_f[11,31] := -0.10893236;
      W_f[11,32] := -0.15593320;
      W_f[11,33] := 0.19035292;
      W_f[11,34] := -0.32335702;
      W_f[11,35] := -0.09812929;
      W_f[11,36] := 0.04003347;
      W_f[11,37] := -0.06675247;
      W_f[11,38] := -0.10143522;
      W_f[11,39] := 0.41168302;
      W_f[12,0] := 0.12018097;
      W_f[12,1] := 0.02609195;
      W_f[12,2] := 0.05892588;
      W_f[12,3] := -0.19573617;
      W_f[12,4] := -0.01478191;
      W_f[12,5] := -0.03957225;
      W_f[12,6] := 0.12785022;
      W_f[12,7] := 0.12322338;
      W_f[12,8] := 0.13078536;
      W_f[12,9] := -0.02882819;
      W_f[12,10] := -0.09103711;
      W_f[12,11] := 0.21010999;
      W_f[12,12] := -0.00687122;
      W_f[12,13] := -0.03154188;
      W_f[12,14] := 0.01292804;
      W_f[12,15] := -0.04617440;
      W_f[12,16] := 0.02552478;
      W_f[12,17] := -0.04503247;
      W_f[12,18] := -0.14453103;
      W_f[12,19] := -0.02086277;
      W_f[12,20] := -0.03427083;
      W_f[12,21] := 0.12834942;
      W_f[12,22] := 0.06980442;
      W_f[12,23] := -0.19849743;
      W_f[12,24] := -0.06221438;
      W_f[12,25] := -0.15592034;
      W_f[12,26] := 0.09680067;
      W_f[12,27] := -0.08721892;
      W_f[12,28] := 0.12007699;
      W_f[12,29] := 0.03281511;
      W_f[12,30] := -0.19682269;
      W_f[12,31] := 0.21656367;
      W_f[12,32] := 0.08357669;
      W_f[12,33] := 0.12308872;
      W_f[12,34] := -0.04732760;
      W_f[12,35] := -0.00432450;
      W_f[12,36] := -0.07603259;
      W_f[12,37] := 0.11208338;
      W_f[12,38] := 0.01071546;
      W_f[12,39] := 0.01300001;
      W_f[13,0] := -0.03169156;
      W_f[13,1] := 0.12357810;
      W_f[13,2] := -0.05470626;
      W_f[13,3] := 0.05454078;
      W_f[13,4] := 0.00082304;
      W_f[13,5] := 0.08142892;
      W_f[13,6] := -0.05739224;
      W_f[13,7] := -0.06891212;
      W_f[13,8] := -0.01340675;
      W_f[13,9] := -0.00828674;
      W_f[13,10] := -0.01201967;
      W_f[13,11] := -0.04392290;
      W_f[13,12] := 0.11794504;
      W_f[13,13] := 0.04059569;
      W_f[13,14] := -0.07634314;
      W_f[13,15] := -0.00757048;
      W_f[13,16] := 0.03631781;
      W_f[13,17] := 0.02680131;
      W_f[13,18] := 0.04420025;
      W_f[13,19] := -0.15575425;
      W_f[13,20] := 0.02057399;
      W_f[13,21] := 0.08036615;
      W_f[13,22] := 0.15103330;
      W_f[13,23] := -0.05069938;
      W_f[13,24] := 0.51470953;
      W_f[13,25] := 0.38624758;
      W_f[13,26] := -0.10547116;
      W_f[13,27] := -0.04113456;
      W_f[13,28] := 0.07717920;
      W_f[13,29] := 0.02030798;
      W_f[13,30] := 0.25870061;
      W_f[13,31] := 0.01822651;
      W_f[13,32] := 0.51183718;
      W_f[13,33] := 0.08568797;
      W_f[13,34] := 0.26839611;
      W_f[13,35] := 0.06110199;
      W_f[13,36] := -0.04498388;
      W_f[13,37] := 0.13735677;
      W_f[13,38] := -0.00712988;
      W_f[13,39] := -0.03385270;
      W_f[14,0] := 0.29193929;
      W_f[14,1] := 0.03370269;
      W_f[14,2] := 0.27688318;
      W_f[14,3] := 0.66428471;
      W_f[14,4] := 0.13141236;
      W_f[14,5] := 0.03623847;
      W_f[14,6] := 0.01996322;
      W_f[14,7] := 0.04668432;
      W_f[14,8] := -0.00427468;
      W_f[14,9] := 0.39187840;
      W_f[14,10] := -0.05717053;
      W_f[14,11] := 0.00223121;
      W_f[14,12] := 0.03597876;
      W_f[14,13] := -0.01569461;
      W_f[14,14] := -0.10418668;
      W_f[14,15] := 0.16508825;
      W_f[14,16] := 0.01595189;
      W_f[14,17] := 0.05152722;
      W_f[14,18] := 0.06324884;
      W_f[14,19] := -0.07842954;
      W_f[14,20] := -0.01252570;
      W_f[14,21] := 0.09333553;
      W_f[14,22] := -0.00592045;
      W_f[14,23] := -0.27803397;
      W_f[14,24] := -0.10406827;
      W_f[14,25] := -0.38742125;
      W_f[14,26] := 0.12681088;
      W_f[14,27] := -0.03332862;
      W_f[14,28] := -0.01383013;
      W_f[14,29] := -0.17758578;
      W_f[14,30] := 0.03754412;
      W_f[14,31] := -0.02210099;
      W_f[14,32] := 0.00901584;
      W_f[14,33] := 0.08400410;
      W_f[14,34] := 0.22526804;
      W_f[14,35] := -0.20718463;
      W_f[14,36] := 0.02469117;
      W_f[14,37] := -0.05200065;
      W_f[14,38] := 0.12603629;
      W_f[14,39] := -0.01085858;
      W_f[15,0] := -0.10406179;
      W_f[15,1] := 0.16952576;
      W_f[15,2] := 0.05386007;
      W_f[15,3] := -0.03501219;
      W_f[15,4] := 0.09106548;
      W_f[15,5] := -0.00729924;
      W_f[15,6] := -0.02398493;
      W_f[15,7] := 0.06805430;
      W_f[15,8] := -0.05002195;
      W_f[15,9] := -0.06974220;
      W_f[15,10] := 0.03180881;
      W_f[15,11] := -0.15035366;
      W_f[15,12] := 0.03008920;
      W_f[15,13] := 0.03584874;
      W_f[15,14] := -0.01684539;
      W_f[15,15] := -0.04871107;
      W_f[15,16] := -0.04879853;
      W_f[15,17] := 0.05787342;
      W_f[15,18] := -0.05507936;
      W_f[15,19] := -0.10834753;
      W_f[15,20] := 0.02284326;
      W_f[15,21] := 0.06631061;
      W_f[15,22] := 0.03862244;
      W_f[15,23] := 0.01920095;
      W_f[15,24] := 0.85719836;
      W_f[15,25] := 0.82220733;
      W_f[15,26] := -0.10065157;
      W_f[15,27] := 0.01829595;
      W_f[15,28] := 0.17395613;
      W_f[15,29] := 0.00457023;
      W_f[15,30] := 0.20811720;
      W_f[15,31] := 0.02074985;
      W_f[15,32] := 0.02153331;
      W_f[15,33] := 0.14867106;
      W_f[15,34] := -0.05699138;
      W_f[15,35] := 0.16990840;
      W_f[15,36] := 0.04588095;
      W_f[15,37] := 0.08796984;
      W_f[15,38] := 0.14537595;
      W_f[15,39] := 0.36507782;
      W_g[0,0] := -0.06437175;
      W_g[0,1] := -0.10304265;
      W_g[0,2] := -0.06360535;
      W_g[0,3] := -0.01407568;
      W_g[0,4] := -0.01109672;
      W_g[0,5] := 0.08344834;
      W_g[0,6] := 0.05906893;
      W_g[0,7] := -0.01122296;
      W_g[0,8] := -0.01076689;
      W_g[0,9] := 0.00505227;
      W_g[0,10] := -0.05708009;
      W_g[0,11] := 0.00101489;
      W_g[0,12] := -0.02898394;
      W_g[0,13] := -0.04387880;
      W_g[0,14] := -0.07387122;
      W_g[0,15] := 0.01959705;
      W_g[0,16] := 0.00128837;
      W_g[0,17] := -0.16131586;
      W_g[0,18] := 0.05533828;
      W_g[0,19] := -0.04145345;
      W_g[0,20] := -0.00717272;
      W_g[0,21] := -0.05831819;
      W_g[0,22] := -0.00424080;
      W_g[0,23] := 0.01501147;
      W_g[0,24] := -0.06262178;
      W_g[0,25] := 0.21272451;
      W_g[0,26] := 0.03131270;
      W_g[0,27] := -0.09072166;
      W_g[0,28] := -0.02835892;
      W_g[0,29] := -0.00038205;
      W_g[0,30] := 0.01341711;
      W_g[0,31] := 0.01420873;
      W_g[0,32] := -0.04364003;
      W_g[0,33] := -0.00602657;
      W_g[0,34] := 0.29625592;
      W_g[0,35] := -0.02899161;
      W_g[0,36] := -0.13954598;
      W_g[0,37] := 0.04718976;
      W_g[0,38] := -0.01878179;
      W_g[0,39] := -0.03507735;
      W_g[1,0] := 0.05452355;
      W_g[1,1] := 0.27387798;
      W_g[1,2] := 0.06841734;
      W_g[1,3] := 0.02098602;
      W_g[1,4] := -0.05067789;
      W_g[1,5] := -0.06117415;
      W_g[1,6] := 0.11808369;
      W_g[1,7] := 0.03169370;
      W_g[1,8] := 0.01715386;
      W_g[1,9] := 0.00421220;
      W_g[1,10] := -0.02094597;
      W_g[1,11] := -0.02231863;
      W_g[1,12] := -0.05272245;
      W_g[1,13] := -0.11053510;
      W_g[1,14] := 0.02985792;
      W_g[1,15] := -0.01159818;
      W_g[1,16] := 0.09040943;
      W_g[1,17] := -0.06152220;
      W_g[1,18] := 0.12156093;
      W_g[1,19] := -0.09465837;
      W_g[1,20] := -0.21014288;
      W_g[1,21] := 0.04188417;
      W_g[1,22] := 0.00875731;
      W_g[1,23] := -0.13488904;
      W_g[1,24] := -0.22675800;
      W_g[1,25] := -0.39127526;
      W_g[1,26] := -0.02196784;
      W_g[1,27] := 0.00777218;
      W_g[1,28] := 0.01569583;
      W_g[1,29] := 0.03508768;
      W_g[1,30] := 0.00428289;
      W_g[1,31] := 0.01024072;
      W_g[1,32] := 0.06771233;
      W_g[1,33] := -0.01064035;
      W_g[1,34] := 0.11919906;
      W_g[1,35] := -0.09515890;
      W_g[1,36] := 0.04105361;
      W_g[1,37] := 0.07846094;
      W_g[1,38] := -0.13942727;
      W_g[1,39] := -0.03954639;
      W_g[2,0] := -0.03289792;
      W_g[2,1] := 0.11950450;
      W_g[2,2] := -0.02634289;
      W_g[2,3] := 0.03330147;
      W_g[2,4] := 0.04832244;
      W_g[2,5] := -0.11697238;
      W_g[2,6] := -0.01332184;
      W_g[2,7] := 0.02626378;
      W_g[2,8] := 0.03550790;
      W_g[2,9] := 0.04916163;
      W_g[2,10] := 0.02250416;
      W_g[2,11] := 0.08283401;
      W_g[2,12] := 0.06788670;
      W_g[2,13] := -0.08117380;
      W_g[2,14] := -0.06664238;
      W_g[2,15] := 0.05342351;
      W_g[2,16] := 0.09484934;
      W_g[2,17] := 0.09736161;
      W_g[2,18] := -0.06697731;
      W_g[2,19] := 0.08243434;
      W_g[2,20] := -0.03165147;
      W_g[2,21] := -0.03695506;
      W_g[2,22] := 0.04532890;
      W_g[2,23] := -0.09410243;
      W_g[2,24] := 0.56509566;
      W_g[2,25] := 0.33052078;
      W_g[2,26] := 0.04841354;
      W_g[2,27] := -0.04202427;
      W_g[2,28] := 0.04029641;
      W_g[2,29] := -0.01918726;
      W_g[2,30] := -0.01533750;
      W_g[2,31] := 0.02825868;
      W_g[2,32] := -0.02275502;
      W_g[2,33] := 0.04718334;
      W_g[2,34] := 0.29532653;
      W_g[2,35] := 0.06282274;
      W_g[2,36] := 0.01098316;
      W_g[2,37] := -0.02031587;
      W_g[2,38] := -0.05517275;
      W_g[2,39] := -0.05778347;
      W_g[3,0] := -0.07797009;
      W_g[3,1] := -0.15111065;
      W_g[3,2] := -0.07784537;
      W_g[3,3] := 0.02676097;
      W_g[3,4] := -0.22783786;
      W_g[3,5] := 0.05178539;
      W_g[3,6] := 0.21769266;
      W_g[3,7] := 0.04195838;
      W_g[3,8] := 0.04416362;
      W_g[3,9] := 0.02287334;
      W_g[3,10] := -0.12170663;
      W_g[3,11] := -0.03924337;
      W_g[3,12] := -0.04121236;
      W_g[3,13] := -0.05717940;
      W_g[3,14] := -0.08332798;
      W_g[3,15] := -0.02212023;
      W_g[3,16] := 0.01032387;
      W_g[3,17] := -0.05978040;
      W_g[3,18] := 0.04619258;
      W_g[3,19] := -0.04743195;
      W_g[3,20] := -0.21954186;
      W_g[3,21] := 0.10694054;
      W_g[3,22] := 0.05955252;
      W_g[3,23] := 0.05258171;
      W_g[3,24] := 0.30032092;
      W_g[3,25] := 0.00568468;
      W_g[3,26] := 0.01930099;
      W_g[3,27] := -0.01615639;
      W_g[3,28] := -0.14664842;
      W_g[3,29] := 0.08185939;
      W_g[3,30] := 0.28245008;
      W_g[3,31] := 0.02146588;
      W_g[3,32] := 0.03048213;
      W_g[3,33] := 0.11187603;
      W_g[3,34] := -0.14845568;
      W_g[3,35] := 0.02283150;
      W_g[3,36] := 0.18844947;
      W_g[3,37] := 0.14089991;
      W_g[3,38] := -0.01001398;
      W_g[3,39] := -0.02703539;
      W_g[4,0] := 0.01343604;
      W_g[4,1] := 0.03630589;
      W_g[4,2] := 0.00586512;
      W_g[4,3] := 0.03330747;
      W_g[4,4] := 0.03309506;
      W_g[4,5] := -0.06498569;
      W_g[4,6] := 0.13742739;
      W_g[4,7] := 0.03903612;
      W_g[4,8] := 0.03540400;
      W_g[4,9] := 0.03336297;
      W_g[4,10] := -0.07885744;
      W_g[4,11] := -0.06243610;
      W_g[4,12] := -0.04985108;
      W_g[4,13] := 0.10830133;
      W_g[4,14] := 0.00163302;
      W_g[4,15] := -0.08075944;
      W_g[4,16] := -0.14402635;
      W_g[4,17] := 0.06278381;
      W_g[4,18] := -0.06662596;
      W_g[4,19] := -0.03559304;
      W_g[4,20] := -0.13648316;
      W_g[4,21] := -0.03422393;
      W_g[4,22] := 0.01963219;
      W_g[4,23] := 0.10719733;
      W_g[4,24] := -0.09623951;
      W_g[4,25] := -0.12038372;
      W_g[4,26] := 0.06311011;
      W_g[4,27] := -0.07769342;
      W_g[4,28] := 0.17828900;
      W_g[4,29] := 0.02263938;
      W_g[4,30] := 0.00952398;
      W_g[4,31] := -0.02689653;
      W_g[4,32] := 0.05671162;
      W_g[4,33] := -0.01929745;
      W_g[4,34] := -0.05658547;
      W_g[4,35] := 0.00156007;
      W_g[4,36] := -0.04812146;
      W_g[4,37] := -0.03719440;
      W_g[4,38] := -0.07058035;
      W_g[4,39] := -0.01562632;
      W_g[5,0] := 0.01347702;
      W_g[5,1] := 0.01319387;
      W_g[5,2] := 0.02702549;
      W_g[5,3] := 0.03099934;
      W_g[5,4] := -0.11858911;
      W_g[5,5] := -0.12051299;
      W_g[5,6] := -0.04255378;
      W_g[5,7] := 0.02337371;
      W_g[5,8] := 0.03234660;
      W_g[5,9] := 0.01507181;
      W_g[5,10] := -0.00441507;
      W_g[5,11] := 0.03045360;
      W_g[5,12] := 0.04173407;
      W_g[5,13] := -0.18411799;
      W_g[5,14] := 0.07539749;
      W_g[5,15] := 0.01865357;
      W_g[5,16] := -0.16913831;
      W_g[5,17] := 0.00040193;
      W_g[5,18] := 0.04012417;
      W_g[5,19] := 0.03515705;
      W_g[5,20] := -0.05170999;
      W_g[5,21] := -0.15163575;
      W_g[5,22] := -0.02755779;
      W_g[5,23] := -0.09758625;
      W_g[5,24] := 0.24352244;
      W_g[5,25] := -0.11935914;
      W_g[5,26] := 0.06693986;
      W_g[5,27] := -0.22207910;
      W_g[5,28] := -0.20637380;
      W_g[5,29] := 0.05818798;
      W_g[5,30] := 0.02412311;
      W_g[5,31] := 0.03364465;
      W_g[5,32] := -0.06383017;
      W_g[5,33] := -0.01355148;
      W_g[5,34] := 0.04340848;
      W_g[5,35] := -0.00615392;
      W_g[5,36] := 0.01951177;
      W_g[5,37] := -0.01499645;
      W_g[5,38] := 0.01239841;
      W_g[5,39] := 0.11211766;
      W_g[6,0] := -0.00913136;
      W_g[6,1] := -0.31391880;
      W_g[6,2] := -0.03205895;
      W_g[6,3] := 0.07225002;
      W_g[6,4] := 0.02337007;
      W_g[6,5] := -0.11176381;
      W_g[6,6] := -0.05067589;
      W_g[6,7] := 0.07076521;
      W_g[6,8] := 0.06279331;
      W_g[6,9] := 0.08101700;
      W_g[6,10] := 0.00219894;
      W_g[6,11] := 0.03236729;
      W_g[6,12] := -0.01466833;
      W_g[6,13] := 0.03211138;
      W_g[6,14] := 0.06749433;
      W_g[6,15] := 0.02329918;
      W_g[6,16] := 0.04367528;
      W_g[6,17] := -0.04910227;
      W_g[6,18] := 0.00852106;
      W_g[6,19] := -0.02368775;
      W_g[6,20] := 0.13064513;
      W_g[6,21] := 0.00328254;
      W_g[6,22] := 0.02020053;
      W_g[6,23] := 0.11741425;
      W_g[6,24] := 0.09362976;
      W_g[6,25] := 0.07101754;
      W_g[6,26] := -0.04242831;
      W_g[6,27] := 0.03521124;
      W_g[6,28] := -0.03469749;
      W_g[6,29] := 0.12673429;
      W_g[6,30] := -0.03175284;
      W_g[6,31] := -0.02456861;
      W_g[6,32] := -0.07071101;
      W_g[6,33] := -0.03622819;
      W_g[6,34] := -0.05097293;
      W_g[6,35] := 0.12351370;
      W_g[6,36] := 0.01210361;
      W_g[6,37] := -0.07118074;
      W_g[6,38] := -0.17139800;
      W_g[6,39] := -0.07202235;
      W_g[7,0] := -0.00221192;
      W_g[7,1] := -0.10343143;
      W_g[7,2] := -0.00175258;
      W_g[7,3] := -0.01847444;
      W_g[7,4] := -0.11821446;
      W_g[7,5] := 0.06384078;
      W_g[7,6] := 0.10368531;
      W_g[7,7] := -0.01418284;
      W_g[7,8] := -0.01802195;
      W_g[7,9] := -0.01371992;
      W_g[7,10] := -0.08365498;
      W_g[7,11] := 0.03279426;
      W_g[7,12] := 0.03902526;
      W_g[7,13] := -0.02570777;
      W_g[7,14] := 0.06307954;
      W_g[7,15] := 0.01467463;
      W_g[7,16] := 0.00880910;
      W_g[7,17] := 0.09958059;
      W_g[7,18] := 0.00496297;
      W_g[7,19] := 0.03075951;
      W_g[7,20] := -0.06976835;
      W_g[7,21] := 0.09910673;
      W_g[7,22] := 0.01788795;
      W_g[7,23] := -0.01338861;
      W_g[7,24] := -0.07418577;
      W_g[7,25] := 0.07377186;
      W_g[7,26] := -0.03523324;
      W_g[7,27] := 0.06126403;
      W_g[7,28] := -0.07607173;
      W_g[7,29] := -0.01105942;
      W_g[7,30] := 0.03793060;
      W_g[7,31] := 0.01525545;
      W_g[7,32] := -0.00270488;
      W_g[7,33] := 0.01759348;
      W_g[7,34] := 0.00930440;
      W_g[7,35] := -0.01158411;
      W_g[7,36] := -0.11851270;
      W_g[7,37] := 0.05517194;
      W_g[7,38] := -0.04390677;
      W_g[7,39] := 0.00916628;
      W_g[8,0] := -0.15320511;
      W_g[8,1] := -0.02698105;
      W_g[8,2] := -0.15616265;
      W_g[8,3] := -0.00037426;
      W_g[8,4] := 0.07145283;
      W_g[8,5] := 0.15556584;
      W_g[8,6] := 0.01163205;
      W_g[8,7] := 0.00025974;
      W_g[8,8] := -0.00305611;
      W_g[8,9] := 0.00339855;
      W_g[8,10] := 0.01435311;
      W_g[8,11] := -0.06739048;
      W_g[8,12] := -0.05513357;
      W_g[8,13] := -0.06115710;
      W_g[8,14] := 0.09001071;
      W_g[8,15] := -0.07062676;
      W_g[8,16] := 0.09425995;
      W_g[8,17] := 0.07710721;
      W_g[8,18] := 0.10256992;
      W_g[8,19] := -0.09351780;
      W_g[8,20] := 0.02987615;
      W_g[8,21] := -0.09316436;
      W_g[8,22] := 0.00862628;
      W_g[8,23] := -0.02039264;
      W_g[8,24] := 0.05032886;
      W_g[8,25] := -0.20768827;
      W_g[8,26] := 0.03280862;
      W_g[8,27] := -0.10336877;
      W_g[8,28] := -0.01109375;
      W_g[8,29] := 0.01177040;
      W_g[8,30] := 0.05040761;
      W_g[8,31] := 0.01287866;
      W_g[8,32] := -0.05836870;
      W_g[8,33] := 0.03837029;
      W_g[8,34] := -0.15856282;
      W_g[8,35] := -0.07470238;
      W_g[8,36] := 0.01450610;
      W_g[8,37] := 0.11253793;
      W_g[8,38] := -0.04236124;
      W_g[8,39] := 0.01533761;
      W_g[9,0] := -0.13535555;
      W_g[9,1] := -0.06505639;
      W_g[9,2] := -0.13579285;
      W_g[9,3] := -0.06444182;
      W_g[9,4] := 0.01908697;
      W_g[9,5] := -0.24531877;
      W_g[9,6] := 0.01296273;
      W_g[9,7] := -0.05682649;
      W_g[9,8] := -0.05677786;
      W_g[9,9] := -0.06395079;
      W_g[9,10] := -0.18071279;
      W_g[9,11] := -0.01403706;
      W_g[9,12] := -0.01820294;
      W_g[9,13] := 0.00699521;
      W_g[9,14] := 0.01161401;
      W_g[9,15] := -0.00308632;
      W_g[9,16] := 0.09676393;
      W_g[9,17] := -0.01729999;
      W_g[9,18] := -0.01128668;
      W_g[9,19] := -0.01986114;
      W_g[9,20] := 0.01903784;
      W_g[9,21] := 0.03708190;
      W_g[9,22] := 0.08796684;
      W_g[9,23] := 0.00702260;
      W_g[9,24] := -0.26771736;
      W_g[9,25] := -0.02212393;
      W_g[9,26] := -0.06138865;
      W_g[9,27] := 0.06166749;
      W_g[9,28] := 0.02480626;
      W_g[9,29] := 0.06521315;
      W_g[9,30] := -0.15108477;
      W_g[9,31] := -0.01764379;
      W_g[9,32] := -0.10532738;
      W_g[9,33] := 0.03247911;
      W_g[9,34] := 0.00060418;
      W_g[9,35] := 0.17793451;
      W_g[9,36] := -0.03480922;
      W_g[9,37] := -0.16084674;
      W_g[9,38] := 0.07908966;
      W_g[9,39] := 0.02495248;
      W_g[10,0] := -0.04868153;
      W_g[10,1] := 0.07170852;
      W_g[10,2] := -0.04725950;
      W_g[10,3] := 0.01684920;
      W_g[10,4] := -0.10642169;
      W_g[10,5] := -0.04727273;
      W_g[10,6] := -0.07462876;
      W_g[10,7] := 0.01728310;
      W_g[10,8] := 0.01981095;
      W_g[10,9] := 0.01254578;
      W_g[10,10] := 0.06902175;
      W_g[10,11] := -0.03850393;
      W_g[10,12] := -0.04260848;
      W_g[10,13] := 0.03856438;
      W_g[10,14] := -0.09470413;
      W_g[10,15] := -0.06301641;
      W_g[10,16] := -0.01483148;
      W_g[10,17] := 0.07461021;
      W_g[10,18] := 0.13068441;
      W_g[10,19] := -0.06515504;
      W_g[10,20] := 0.08656729;
      W_g[10,21] := 0.02321765;
      W_g[10,22] := -0.00932684;
      W_g[10,23] := 0.05053019;
      W_g[10,24] := 0.12723380;
      W_g[10,25] := 0.13141626;
      W_g[10,26] := -0.03516380;
      W_g[10,27] := 0.02526680;
      W_g[10,28] := -0.18210968;
      W_g[10,29] := -0.04132932;
      W_g[10,30] := 0.01944728;
      W_g[10,31] := 0.01472420;
      W_g[10,32] := -0.03706682;
      W_g[10,33] := 0.01090265;
      W_g[10,34] := 0.17765786;
      W_g[10,35] := -0.01664727;
      W_g[10,36] := -0.05660886;
      W_g[10,37] := 0.03716451;
      W_g[10,38] := -0.01593407;
      W_g[10,39] := -0.05980631;
      W_g[11,0] := -0.07778873;
      W_g[11,1] := 0.13476834;
      W_g[11,2] := -0.07938315;
      W_g[11,3] := 0.05070763;
      W_g[11,4] := -0.00296141;
      W_g[11,5] := -0.03763780;
      W_g[11,6] := 0.01238506;
      W_g[11,7] := 0.06416834;
      W_g[11,8] := 0.04759337;
      W_g[11,9] := 0.05471492;
      W_g[11,10] := 0.05613361;
      W_g[11,11] := -0.03514048;
      W_g[11,12] := 0.00023959;
      W_g[11,13] := 0.07004435;
      W_g[11,14] := 0.13153584;
      W_g[11,15] := 0.00372343;
      W_g[11,16] := 0.00074738;
      W_g[11,17] := -0.11343645;
      W_g[11,18] := 0.00006006;
      W_g[11,19] := -0.01685918;
      W_g[11,20] := 0.01445182;
      W_g[11,21] := 0.06210520;
      W_g[11,22] := 0.02249984;
      W_g[11,23] := 0.07355771;
      W_g[11,24] := 0.31212780;
      W_g[11,25] := 0.28221378;
      W_g[11,26] := -0.00655897;
      W_g[11,27] := 0.09088862;
      W_g[11,28] := 0.03146487;
      W_g[11,29] := -0.02166439;
      W_g[11,30] := -0.00286892;
      W_g[11,31] := 0.01861817;
      W_g[11,32] := -0.02104462;
      W_g[11,33] := 0.05356301;
      W_g[11,34] := 0.22107139;
      W_g[11,35] := 0.08230665;
      W_g[11,36] := -0.04974785;
      W_g[11,37] := 0.02396704;
      W_g[11,38] := 0.02959024;
      W_g[11,39] := 0.16378370;
      W_g[12,0] := -0.05897811;
      W_g[12,1] := 0.04489198;
      W_g[12,2] := -0.05050897;
      W_g[12,3] := 0.00414122;
      W_g[12,4] := -0.12534045;
      W_g[12,5] := 0.01220162;
      W_g[12,6] := -0.07195626;
      W_g[12,7] := -0.00308424;
      W_g[12,8] := 0.00341901;
      W_g[12,9] := -0.00221285;
      W_g[12,10] := 0.05365397;
      W_g[12,11] := -0.07171583;
      W_g[12,12] := -0.07715646;
      W_g[12,13] := -0.15127288;
      W_g[12,14] := 0.01169638;
      W_g[12,15] := -0.05661723;
      W_g[12,16] := 0.02522748;
      W_g[12,17] := -0.03785696;
      W_g[12,18] := -0.64070398;
      W_g[12,19] := -0.05478346;
      W_g[12,20] := 0.01582275;
      W_g[12,21] := 0.00480355;
      W_g[12,22] := -0.12825850;
      W_g[12,23] := -0.11299890;
      W_g[12,24] := 0.05207260;
      W_g[12,25] := 0.01753274;
      W_g[12,26] := -0.00488592;
      W_g[12,27] := -0.02255455;
      W_g[12,28] := -0.19238769;
      W_g[12,29] := 0.01013393;
      W_g[12,30] := 0.02022840;
      W_g[12,31] := 0.00866093;
      W_g[12,32] := -0.15646824;
      W_g[12,33] := 0.03487159;
      W_g[12,34] := -0.02648159;
      W_g[12,35] := -0.01117676;
      W_g[12,36] := -0.02055392;
      W_g[12,37] := -0.04472685;
      W_g[12,38] := -0.11415342;
      W_g[12,39] := -0.02697767;
      W_g[13,0] := 0.05595589;
      W_g[13,1] := -0.07274999;
      W_g[13,2] := 0.05476713;
      W_g[13,3] := 0.03637930;
      W_g[13,4] := -0.14596705;
      W_g[13,5] := -0.07975005;
      W_g[13,6] := 0.03538230;
      W_g[13,7] := 0.04020952;
      W_g[13,8] := 0.04126918;
      W_g[13,9] := 0.04235730;
      W_g[13,10] := -0.02485134;
      W_g[13,11] := 0.02735355;
      W_g[13,12] := 0.01234699;
      W_g[13,13] := 0.03710405;
      W_g[13,14] := -0.01809123;
      W_g[13,15] := 0.03689704;
      W_g[13,16] := 0.20435552;
      W_g[13,17] := 0.00377080;
      W_g[13,18] := -0.03157456;
      W_g[13,19] := 0.01731828;
      W_g[13,20] := -0.06259499;
      W_g[13,21] := -0.06937376;
      W_g[13,22] := -0.04025269;
      W_g[13,23] := 0.10691475;
      W_g[13,24] := 0.15896399;
      W_g[13,25] := -0.04750140;
      W_g[13,26] := 0.04742527;
      W_g[13,27] := -0.10945089;
      W_g[13,28] := -0.11246481;
      W_g[13,29] := 0.02072454;
      W_g[13,30] := -0.04956476;
      W_g[13,31] := -0.01100769;
      W_g[13,32] := -0.04496330;
      W_g[13,33] := -0.07340268;
      W_g[13,34] := 0.09542960;
      W_g[13,35] := -0.06956401;
      W_g[13,36] := -0.05015138;
      W_g[13,37] := -0.01480982;
      W_g[13,38] := 0.04396211;
      W_g[13,39] := 0.00700256;
      W_g[14,0] := 0.08032657;
      W_g[14,1] := 0.17840010;
      W_g[14,2] := 0.07731044;
      W_g[14,3] := -0.09140022;
      W_g[14,4] := -0.08219359;
      W_g[14,5] := 0.05311288;
      W_g[14,6] := -0.03072528;
      W_g[14,7] := -0.12227103;
      W_g[14,8] := -0.10546146;
      W_g[14,9] := -0.12072457;
      W_g[14,10] := -0.09533292;
      W_g[14,11] := -0.00337938;
      W_g[14,12] := 0.01313734;
      W_g[14,13] := 0.16531847;
      W_g[14,14] := 0.07715569;
      W_g[14,15] := 0.02926527;
      W_g[14,16] := 0.01751664;
      W_g[14,17] := -0.03058667;
      W_g[14,18] := -0.25051984;
      W_g[14,19] := -0.00634941;
      W_g[14,20] := -0.03018456;
      W_g[14,21] := -0.05928081;
      W_g[14,22] := 0.05027040;
      W_g[14,23] := 0.09324472;
      W_g[14,24] := -0.22232357;
      W_g[14,25] := 0.20548849;
      W_g[14,26] := 0.04399953;
      W_g[14,27] := -0.08267367;
      W_g[14,28] := -0.03239481;
      W_g[14,29] := 0.00585578;
      W_g[14,30] := 0.03364217;
      W_g[14,31] := 0.01409262;
      W_g[14,32] := 0.09821244;
      W_g[14,33] := 0.08529360;
      W_g[14,34] := -0.15575923;
      W_g[14,35] := -0.00937407;
      W_g[14,36] := 0.05313390;
      W_g[14,37] := -0.00805885;
      W_g[14,38] := -0.15908019;
      W_g[14,39] := -0.07129225;
      W_g[15,0] := 0.14802523;
      W_g[15,1] := -0.09804792;
      W_g[15,2] := 0.14636119;
      W_g[15,3] := -0.02253639;
      W_g[15,4] := 0.06714331;
      W_g[15,5] := -0.07940288;
      W_g[15,6] := -0.02956429;
      W_g[15,7] := -0.02010203;
      W_g[15,8] := -0.02122243;
      W_g[15,9] := -0.00691266;
      W_g[15,10] := -0.03708303;
      W_g[15,11] := -0.10704023;
      W_g[15,12] := -0.11317661;
      W_g[15,13] := -0.00916757;
      W_g[15,14] := -0.00417171;
      W_g[15,15] := -0.09912409;
      W_g[15,16] := 0.05694117;
      W_g[15,17] := -0.00757575;
      W_g[15,18] := 0.01970402;
      W_g[15,19] := -0.11384802;
      W_g[15,20] := 0.04223837;
      W_g[15,21] := 0.00676507;
      W_g[15,22] := 0.07206889;
      W_g[15,23] := -0.02210784;
      W_g[15,24] := 0.33264917;
      W_g[15,25] := 0.19025688;
      W_g[15,26] := 0.00426384;
      W_g[15,27] := -0.00031623;
      W_g[15,28] := 0.02923820;
      W_g[15,29] := -0.13043131;
      W_g[15,30] := 0.01179718;
      W_g[15,31] := 0.02720840;
      W_g[15,32] := 0.16045739;
      W_g[15,33] := -0.03539550;
      W_g[15,34] := 0.02744242;
      W_g[15,35] := 0.05568860;
      W_g[15,36] := -0.06267934;
      W_g[15,37] := -0.07925017;
      W_g[15,38] := 0.03805197;
      W_g[15,39] := -0.00476847;
      W_o[0,0] := 0.03012275;
      W_o[0,1] := -0.06497240;
      W_o[0,2] := -0.21605290;
      W_o[0,3] := -0.19879378;
      W_o[0,4] := 0.25872990;
      W_o[0,5] := -0.12768269;
      W_o[0,6] := 0.28797144;
      W_o[0,7] := -0.07324373;
      W_o[0,8] := -0.08770406;
      W_o[0,9] := 0.12128527;
      W_o[0,10] := -0.30661353;
      W_o[0,11] := -0.83766937;
      W_o[0,12] := 0.08383763;
      W_o[0,13] := 0.06981274;
      W_o[0,14] := -0.19680905;
      W_o[0,15] := -0.38373759;
      W_o[0,16] := -0.28850493;
      W_o[0,17] := -0.42365679;
      W_o[0,18] := 0.36578110;
      W_o[0,19] := -0.00007986;
      W_o[0,20] := -0.30372488;
      W_o[0,21] := -0.00331270;
      W_o[0,22] := 0.90026724;
      W_o[0,23] := -0.37525588;
      W_o[0,24] := 1.50997412;
      W_o[0,25] := 1.66138411;
      W_o[0,26] := -0.48010135;
      W_o[0,27] := -0.17736135;
      W_o[0,28] := -0.29523391;
      W_o[0,29] := -0.71863556;
      W_o[0,30] := 0.54567719;
      W_o[0,31] := 0.16052328;
      W_o[0,32] := 0.56617969;
      W_o[0,33] := 0.54288220;
      W_o[0,34] := 1.32341599;
      W_o[0,35] := 0.68102258;
      W_o[0,36] := 0.27216136;
      W_o[0,37] := 0.60816181;
      W_o[0,38] := 0.13368255;
      W_o[0,39] := 0.21520153;
      W_o[1,0] := 0.47674629;
      W_o[1,1] := 0.15082929;
      W_o[1,2] := 0.11851368;
      W_o[1,3] := -0.17266349;
      W_o[1,4] := 0.26910278;
      W_o[1,5] := -0.03040568;
      W_o[1,6] := 0.33718312;
      W_o[1,7] := 0.21070869;
      W_o[1,8] := 0.32091576;
      W_o[1,9] := -0.01046208;
      W_o[1,10] := -0.14176907;
      W_o[1,11] := -0.11895081;
      W_o[1,12] := 0.17483769;
      W_o[1,13] := -0.24414009;
      W_o[1,14] := 0.00898027;
      W_o[1,15] := -0.11913206;
      W_o[1,16] := -0.17226383;
      W_o[1,17] := -0.03561071;
      W_o[1,18] := 0.80387825;
      W_o[1,19] := 0.09534956;
      W_o[1,20] := -0.34201932;
      W_o[1,21] := 0.45919308;
      W_o[1,22] := 0.22873488;
      W_o[1,23] := -0.20797899;
      W_o[1,24] := 0.11995200;
      W_o[1,25] := 0.03844377;
      W_o[1,26] := -0.11905818;
      W_o[1,27] := -0.10153977;
      W_o[1,28] := 0.21479538;
      W_o[1,29] := -0.06160569;
      W_o[1,30] := 0.03565846;
      W_o[1,31] := 0.02235219;
      W_o[1,32] := 0.14506997;
      W_o[1,33] := 0.11349452;
      W_o[1,34] := -0.05920382;
      W_o[1,35] := -0.22101414;
      W_o[1,36] := -0.05821102;
      W_o[1,37] := 0.01527586;
      W_o[1,38] := 0.33995131;
      W_o[1,39] := -0.08461418;
      W_o[2,0] := -0.04041630;
      W_o[2,1] := 0.24293591;
      W_o[2,2] := -0.08497260;
      W_o[2,3] := 0.00539105;
      W_o[2,4] := 0.23852527;
      W_o[2,5] := 0.47765291;
      W_o[2,6] := 0.03909414;
      W_o[2,7] := 0.18794830;
      W_o[2,8] := 0.13327233;
      W_o[2,9] := 0.07918805;
      W_o[2,10] := 0.26217058;
      W_o[2,11] := -0.40030104;
      W_o[2,12] := -0.32532111;
      W_o[2,13] := -0.16847309;
      W_o[2,14] := 0.05510291;
      W_o[2,15] := -0.21259028;
      W_o[2,16] := 0.15200765;
      W_o[2,17] := 0.06253191;
      W_o[2,18] := -0.29971015;
      W_o[2,19] := -0.37370089;
      W_o[2,20] := -0.09585105;
      W_o[2,21] := 0.00693277;
      W_o[2,22] := 0.11310136;
      W_o[2,23] := 0.00886431;
      W_o[2,24] := -0.06598823;
      W_o[2,25] := -0.13190241;
      W_o[2,26] := -0.02707478;
      W_o[2,27] := -0.04556934;
      W_o[2,28] := 0.26014969;
      W_o[2,29] := 0.01684864;
      W_o[2,30] := 0.13470268;
      W_o[2,31] := 0.05851230;
      W_o[2,32] := -0.12677705;
      W_o[2,33] := -0.01981959;
      W_o[2,34] := -0.17276917;
      W_o[2,35] := -0.16546290;
      W_o[2,36] := -0.10995308;
      W_o[2,37] := -0.18001004;
      W_o[2,38] := -0.24247925;
      W_o[2,39] := 0.61191142;
      W_o[3,0] := 0.16471930;
      W_o[3,1] := 0.11132648;
      W_o[3,2] := -0.31437626;
      W_o[3,3] := -0.00312838;
      W_o[3,4] := 0.15883976;
      W_o[3,5] := 0.13949926;
      W_o[3,6] := 0.08379781;
      W_o[3,7] := 0.33693710;
      W_o[3,8] := 0.06524722;
      W_o[3,9] := 0.07056973;
      W_o[3,10] := -0.06616178;
      W_o[3,11] := -0.16736726;
      W_o[3,12] := 0.08917592;
      W_o[3,13] := -0.17018434;
      W_o[3,14] := -0.18161288;
      W_o[3,15] := -0.15950353;
      W_o[3,16] := 0.03381697;
      W_o[3,17] := -0.10723723;
      W_o[3,18] := 0.12991950;
      W_o[3,19] := -0.24874295;
      W_o[3,20] := -0.16043054;
      W_o[3,21] := 0.05139644;
      W_o[3,22] := -0.21882506;
      W_o[3,23] := -0.18416485;
      W_o[3,24] := 0.07846256;
      W_o[3,25] := -0.11334875;
      W_o[3,26] := 0.12250697;
      W_o[3,27] := -0.28703529;
      W_o[3,28] := 0.01738480;
      W_o[3,29] := 0.16785549;
      W_o[3,30] := -0.36865276;
      W_o[3,31] := -0.13739067;
      W_o[3,32] := -0.29462498;
      W_o[3,33] := 0.21976557;
      W_o[3,34] := -0.07948454;
      W_o[3,35] := 0.02594316;
      W_o[3,36] := 0.05661822;
      W_o[3,37] := 0.01088546;
      W_o[3,38] := -0.08284936;
      W_o[3,39] := -0.04624766;
      W_o[4,0] := -0.14103185;
      W_o[4,1] := 0.08273518;
      W_o[4,2] := 0.22572006;
      W_o[4,3] := -0.09172086;
      W_o[4,4] := -0.11351925;
      W_o[4,5] := -0.11563966;
      W_o[4,6] := -0.02519809;
      W_o[4,7] := -0.07279444;
      W_o[4,8] := -0.02726443;
      W_o[4,9] := 0.24529301;
      W_o[4,10] := 0.00560312;
      W_o[4,11] := -0.10246013;
      W_o[4,12] := -0.01757793;
      W_o[4,13] := -0.24487424;
      W_o[4,14] := -0.06368216;
      W_o[4,15] := -0.13879970;
      W_o[4,16] := -0.44478709;
      W_o[4,17] := 0.04339453;
      W_o[4,18] := 0.16379321;
      W_o[4,19] := -0.20043707;
      W_o[4,20] := 0.42696035;
      W_o[4,21] := 0.27584559;
      W_o[4,22] := 0.03638229;
      W_o[4,23] := -0.27982605;
      W_o[4,24] := 0.89867461;
      W_o[4,25] := 1.06885791;
      W_o[4,26] := -0.18278535;
      W_o[4,27] := 0.10765752;
      W_o[4,28] := -0.34283939;
      W_o[4,29] := -0.11070991;
      W_o[4,30] := 0.22111182;
      W_o[4,31] := 0.08323267;
      W_o[4,32] := -0.01194908;
      W_o[4,33] := 0.12561017;
      W_o[4,34] := 0.34231696;
      W_o[4,35] := 0.13452707;
      W_o[4,36] := 0.03836655;
      W_o[4,37] := 0.23499574;
      W_o[4,38] := 0.10191178;
      W_o[4,39] := -0.01685481;
      W_o[5,0] := 0.00612297;
      W_o[5,1] := 0.16049230;
      W_o[5,2] := 0.05772954;
      W_o[5,3] := 0.30941138;
      W_o[5,4] := 0.33486956;
      W_o[5,5] := 0.49437922;
      W_o[5,6] := 0.32231948;
      W_o[5,7] := -0.08946527;
      W_o[5,8] := 0.05433865;
      W_o[5,9] := 0.08644859;
      W_o[5,10] := 0.03819366;
      W_o[5,11] := -0.25630406;
      W_o[5,12] := 0.03281128;
      W_o[5,13] := 0.10912674;
      W_o[5,14] := 0.42209649;
      W_o[5,15] := -0.20385981;
      W_o[5,16] := 0.13880774;
      W_o[5,17] := 0.05286700;
      W_o[5,18] := 0.50802064;
      W_o[5,19] := 0.05522392;
      W_o[5,20] := 0.01618003;
      W_o[5,21] := 0.24978748;
      W_o[5,22] := 0.45558840;
      W_o[5,23] := -0.45151913;
      W_o[5,24] := 1.27194798;
      W_o[5,25] := 1.37390590;
      W_o[5,26] := -0.17285615;
      W_o[5,27] := -0.16947708;
      W_o[5,28] := 0.03011410;
      W_o[5,29] := -0.07647764;
      W_o[5,30] := 0.32299334;
      W_o[5,31] := -0.05761106;
      W_o[5,32] := -0.03715022;
      W_o[5,33] := -0.08140672;
      W_o[5,34] := 0.70606804;
      W_o[5,35] := 0.06046238;
      W_o[5,36] := 0.09497046;
      W_o[5,37] := 0.00204190;
      W_o[5,38] := 0.35044545;
      W_o[5,39] := -0.03814309;
      W_o[6,0] := 0.21213289;
      W_o[6,1] := 0.38289395;
      W_o[6,2] := 0.17430520;
      W_o[6,3] := 0.11534344;
      W_o[6,4] := -0.24694002;
      W_o[6,5] := 0.17775424;
      W_o[6,6] := -0.03827825;
      W_o[6,7] := 0.12728505;
      W_o[6,8] := 0.02084523;
      W_o[6,9] := 0.59846830;
      W_o[6,10] := 0.57359946;
      W_o[6,11] := 0.01237764;
      W_o[6,12] := -0.23363464;
      W_o[6,13] := -0.28108862;
      W_o[6,14] := -0.00023332;
      W_o[6,15] := 0.05771344;
      W_o[6,16] := -0.10366344;
      W_o[6,17] := 0.15887503;
      W_o[6,18] := 0.36715120;
      W_o[6,19] := 0.02018637;
      W_o[6,20] := -0.67914212;
      W_o[6,21] := -0.28104323;
      W_o[6,22] := 0.12654921;
      W_o[6,23] := -0.62203121;
      W_o[6,24] := 1.59809518;
      W_o[6,25] := 1.52839673;
      W_o[6,26] := -0.17257482;
      W_o[6,27] := 0.03214070;
      W_o[6,28] := 0.17203955;
      W_o[6,29] := -0.01515619;
      W_o[6,30] := 0.09394256;
      W_o[6,31] := -0.26124841;
      W_o[6,32] := -0.15100044;
      W_o[6,33] := -0.18846129;
      W_o[6,34] := 0.43594933;
      W_o[6,35] := -0.46914530;
      W_o[6,36] := 0.08818512;
      W_o[6,37] := -0.21027035;
      W_o[6,38] := 0.51119655;
      W_o[6,39] := 0.21959713;
      W_o[7,0] := 0.00880489;
      W_o[7,1] := 0.16389218;
      W_o[7,2] := -0.27187598;
      W_o[7,3] := -0.08521115;
      W_o[7,4] := -0.23227458;
      W_o[7,5] := 0.18615586;
      W_o[7,6] := 0.39290863;
      W_o[7,7] := 0.24668033;
      W_o[7,8] := -0.07169566;
      W_o[7,9] := 0.02574087;
      W_o[7,10] := -0.06324504;
      W_o[7,11] := -0.67390841;
      W_o[7,12] := -0.37920567;
      W_o[7,13] := -0.04154281;
      W_o[7,14] := -0.22709990;
      W_o[7,15] := -0.51499224;
      W_o[7,16] := 0.55693632;
      W_o[7,17] := 0.17397258;
      W_o[7,18] := 0.24895263;
      W_o[7,19] := -0.35976043;
      W_o[7,20] := 0.16014469;
      W_o[7,21] := 0.00632684;
      W_o[7,22] := 0.58045584;
      W_o[7,23] := -0.18180482;
      W_o[7,24] := 0.63141513;
      W_o[7,25] := 0.71103871;
      W_o[7,26] := 0.01249222;
      W_o[7,27] := -0.08925499;
      W_o[7,28] := 0.34805465;
      W_o[7,29] := -0.45465195;
      W_o[7,30] := 0.62483996;
      W_o[7,31] := 0.14616422;
      W_o[7,32] := 0.31024432;
      W_o[7,33] := 0.07542430;
      W_o[7,34] := 0.75282276;
      W_o[7,35] := 0.12564446;
      W_o[7,36] := -0.13589483;
      W_o[7,37] := 0.48068321;
      W_o[7,38] := 0.04344949;
      W_o[7,39] := 0.02534149;
      W_o[8,0] := -0.04438690;
      W_o[8,1] := 0.03676237;
      W_o[8,2] := -0.19825736;
      W_o[8,3] := -0.25087598;
      W_o[8,4] := -0.04120675;
      W_o[8,5] := -0.06573436;
      W_o[8,6] := 0.02562640;
      W_o[8,7] := -0.20834209;
      W_o[8,8] := 0.00342313;
      W_o[8,9] := -0.03044749;
      W_o[8,10] := -0.20552474;
      W_o[8,11] := -0.34068409;
      W_o[8,12] := 0.04947798;
      W_o[8,13] := -0.27354696;
      W_o[8,14] := -0.03973003;
      W_o[8,15] := -0.06131041;
      W_o[8,16] := 0.39990726;
      W_o[8,17] := -0.00424056;
      W_o[8,18] := 0.03408558;
      W_o[8,19] := -0.29740992;
      W_o[8,20] := -0.15217216;
      W_o[8,21] := 0.26448521;
      W_o[8,22] := 0.29771900;
      W_o[8,23] := -0.22402741;
      W_o[8,24] := 0.62246871;
      W_o[8,25] := 0.40032035;
      W_o[8,26] := -0.18099377;
      W_o[8,27] := 0.00593790;
      W_o[8,28] := -0.03178592;
      W_o[8,29] := 0.13063684;
      W_o[8,30] := 0.06884465;
      W_o[8,31] := 0.20790291;
      W_o[8,32] := 0.30237511;
      W_o[8,33] := 0.22670560;
      W_o[8,34] := 0.28230992;
      W_o[8,35] := -0.14857355;
      W_o[8,36] := 0.02271347;
      W_o[8,37] := -0.11579860;
      W_o[8,38] := 0.25802994;
      W_o[8,39] := 0.22013596;
      W_o[9,0] := -0.31326410;
      W_o[9,1] := -0.06183321;
      W_o[9,2] := -0.11908967;
      W_o[9,3] := -0.14727123;
      W_o[9,4] := -0.20513229;
      W_o[9,5] := -0.61921901;
      W_o[9,6] := 0.13875237;
      W_o[9,7] := -0.31663069;
      W_o[9,8] := -0.95899773;
      W_o[9,9] := 0.07396720;
      W_o[9,10] := -0.33321306;
      W_o[9,11] := 0.07539017;
      W_o[9,12] := 0.04058671;
      W_o[9,13] := -0.03272064;
      W_o[9,14] := 0.00082348;
      W_o[9,15] := 0.03252422;
      W_o[9,16] := -0.18708903;
      W_o[9,17] := 0.03206202;
      W_o[9,18] := -0.11099736;
      W_o[9,19] := -0.20952043;
      W_o[9,20] := -0.51351130;
      W_o[9,21] := 0.19206487;
      W_o[9,22] := -0.01424127;
      W_o[9,23] := -0.00173319;
      W_o[9,24] := -0.08532184;
      W_o[9,25] := -0.28213185;
      W_o[9,26] := -0.03178848;
      W_o[9,27] := -0.05777990;
      W_o[9,28] := 0.23150153;
      W_o[9,29] := 0.07085361;
      W_o[9,30] := 0.19510473;
      W_o[9,31] := 0.08876722;
      W_o[9,32] := 0.14023726;
      W_o[9,33] := 0.28219888;
      W_o[9,34] := 0.16065253;
      W_o[9,35] := -0.19289231;
      W_o[9,36] := 0.01568728;
      W_o[9,37] := -0.18600458;
      W_o[9,38] := 0.09268271;
      W_o[9,39] := -0.01587286;
      W_o[10,0] := -0.02192705;
      W_o[10,1] := 0.23295419;
      W_o[10,2] := -0.00188665;
      W_o[10,3] := 0.14379205;
      W_o[10,4] := 0.25322789;
      W_o[10,5] := 0.45421651;
      W_o[10,6] := 0.32603258;
      W_o[10,7] := 0.12987848;
      W_o[10,8] := -0.03717055;
      W_o[10,9] := 0.06002445;
      W_o[10,10] := -0.01521991;
      W_o[10,11] := -0.31102183;
      W_o[10,12] := -0.20097059;
      W_o[10,13] := 0.05733368;
      W_o[10,14] := -0.34040114;
      W_o[10,15] := -0.47372326;
      W_o[10,16] := 0.03586001;
      W_o[10,17] := 0.12237096;
      W_o[10,18] := 0.30013287;
      W_o[10,19] := -0.05952299;
      W_o[10,20] := -0.12228516;
      W_o[10,21] := 0.16445750;
      W_o[10,22] := 0.35036501;
      W_o[10,23] := -0.32127064;
      W_o[10,24] := 1.07512653;
      W_o[10,25] := 1.03137481;
      W_o[10,26] := -0.08657660;
      W_o[10,27] := -0.34745640;
      W_o[10,28] := 0.09863426;
      W_o[10,29] := -0.21327834;
      W_o[10,30] := 0.38512465;
      W_o[10,31] := 0.11822507;
      W_o[10,32] := 0.34400395;
      W_o[10,33] := 0.38991973;
      W_o[10,34] := 0.73926532;
      W_o[10,35] := 0.20041491;
      W_o[10,36] := -0.05608039;
      W_o[10,37] := 0.22759920;
      W_o[10,38] := -0.04267087;
      W_o[10,39] := 0.28368264;
      W_o[11,0] := -0.18096527;
      W_o[11,1] := 0.10150715;
      W_o[11,2] := -0.13597865;
      W_o[11,3] := -0.33922195;
      W_o[11,4] := 0.01738593;
      W_o[11,5] := 0.00192241;
      W_o[11,6] := -0.02194121;
      W_o[11,7] := -0.15470769;
      W_o[11,8] := 0.06660517;
      W_o[11,9] := -0.13483830;
      W_o[11,10] := -0.13476704;
      W_o[11,11] := -0.17826928;
      W_o[11,12] := 0.14727013;
      W_o[11,13] := -0.27866167;
      W_o[11,14] := 0.09056337;
      W_o[11,15] := -0.07600223;
      W_o[11,16] := 0.04268850;
      W_o[11,17] := 0.19397056;
      W_o[11,18] := 0.06352299;
      W_o[11,19] := -0.31846920;
      W_o[11,20] := -0.08175273;
      W_o[11,21] := 0.15625605;
      W_o[11,22] := -0.13186333;
      W_o[11,23] := -0.42270559;
      W_o[11,24] := 0.03163491;
      W_o[11,25] := 0.30734661;
      W_o[11,26] := 0.18475358;
      W_o[11,27] := -0.19691366;
      W_o[11,28] := 0.12857850;
      W_o[11,29] := 0.02137278;
      W_o[11,30] := -0.08936202;
      W_o[11,31] := 0.27817145;
      W_o[11,32] := -0.09503862;
      W_o[11,33] := -0.16586573;
      W_o[11,34] := -0.12783831;
      W_o[11,35] := -0.16244578;
      W_o[11,36] := 0.19029213;
      W_o[11,37] := 0.12786503;
      W_o[11,38] := -0.07075812;
      W_o[11,39] := 0.42838198;
      W_o[12,0] := -0.12199911;
      W_o[12,1] := 0.03823468;
      W_o[12,2] := 0.01577434;
      W_o[12,3] := 0.14700466;
      W_o[12,4] := 0.07602670;
      W_o[12,5] := -0.05943288;
      W_o[12,6] := 0.12184242;
      W_o[12,7] := -0.40920180;
      W_o[12,8] := -0.01477545;
      W_o[12,9] := 0.10503855;
      W_o[12,10] := -0.06524223;
      W_o[12,11] := -0.04999274;
      W_o[12,12] := 0.35217780;
      W_o[12,13] := -0.07877419;
      W_o[12,14] := 0.09900068;
      W_o[12,15] := 0.05063246;
      W_o[12,16] := 0.10215761;
      W_o[12,17] := -0.11722887;
      W_o[12,18] := 0.07565860;
      W_o[12,19] := -0.08223618;
      W_o[12,20] := -0.28514686;
      W_o[12,21] := -0.00324072;
      W_o[12,22] := 0.06362450;
      W_o[12,23] := -0.18293576;
      W_o[12,24] := -0.30758157;
      W_o[12,25] := -0.27201420;
      W_o[12,26] := 0.16889216;
      W_o[12,27] := 0.06790268;
      W_o[12,28] := 0.09229479;
      W_o[12,29] := -0.02702256;
      W_o[12,30] := 0.04384379;
      W_o[12,31] := -0.27102986;
      W_o[12,32] := -0.19300066;
      W_o[12,33] := 0.32361642;
      W_o[12,34] := 0.00694379;
      W_o[12,35] := 0.05657077;
      W_o[12,36] := -0.12715450;
      W_o[12,37] := -0.12429225;
      W_o[12,38] := 0.28967735;
      W_o[12,39] := -0.08116662;
      W_o[13,0] := 0.36894697;
      W_o[13,1] := 0.11307722;
      W_o[13,2] := 0.54710245;
      W_o[13,3] := -0.38298383;
      W_o[13,4] := 0.64984828;
      W_o[13,5] := -0.26027730;
      W_o[13,6] := 0.20946513;
      W_o[13,7] := 0.02607361;
      W_o[13,8] := -0.11126383;
      W_o[13,9] := -0.06411502;
      W_o[13,10] := -0.03624791;
      W_o[13,11] := -0.04085876;
      W_o[13,12] := -0.34974921;
      W_o[13,13] := -0.16055733;
      W_o[13,14] := 0.17827825;
      W_o[13,15] := -0.04494572;
      W_o[13,16] := 0.14996555;
      W_o[13,17] := -0.11093142;
      W_o[13,18] := 0.53310508;
      W_o[13,19] := -0.44423905;
      W_o[13,20] := -0.07231531;
      W_o[13,21] := 0.36429852;
      W_o[13,22] := 0.57765251;
      W_o[13,23] := -0.14467408;
      W_o[13,24] := 1.53784323;
      W_o[13,25] := 1.40646410;
      W_o[13,26] := -0.19820833;
      W_o[13,27] := 0.25259751;
      W_o[13,28] := 0.10905714;
      W_o[13,29] := -0.38636085;
      W_o[13,30] := 0.31986794;
      W_o[13,31] := -0.06557760;
      W_o[13,32] := 0.15913956;
      W_o[13,33] := 0.33023718;
      W_o[13,34] := 0.80108660;
      W_o[13,35] := 0.00219575;
      W_o[13,36] := 0.31940156;
      W_o[13,37] := 0.32923642;
      W_o[13,38] := 0.28953710;
      W_o[13,39] := 0.14381041;
      W_o[14,0] := -0.06043304;
      W_o[14,1] := 0.14638376;
      W_o[14,2] := 0.18131150;
      W_o[14,3] := -0.44611737;
      W_o[14,4] := -0.08022243;
      W_o[14,5] := 0.12152494;
      W_o[14,6] := -0.09096271;
      W_o[14,7] := -0.08817829;
      W_o[14,8] := -0.41048923;
      W_o[14,9] := 0.00550563;
      W_o[14,10] := 0.02338252;
      W_o[14,11] := 0.03576816;
      W_o[14,12] := 0.09025624;
      W_o[14,13] := -0.16595198;
      W_o[14,14] := -0.18596272;
      W_o[14,15] := -0.09394215;
      W_o[14,16] := -0.06208068;
      W_o[14,17] := -0.00717838;
      W_o[14,18] := 0.19969238;
      W_o[14,19] := 0.01073706;
      W_o[14,20] := -0.18231358;
      W_o[14,21] := 0.01420894;
      W_o[14,22] := -0.10174545;
      W_o[14,23] := -0.49757239;
      W_o[14,24] := -0.46729681;
      W_o[14,25] := -0.29240492;
      W_o[14,26] := -0.19052799;
      W_o[14,27] := -0.16709423;
      W_o[14,28] := -0.01935058;
      W_o[14,29] := -0.14249825;
      W_o[14,30] := -0.15881291;
      W_o[14,31] := 0.20393510;
      W_o[14,32] := -0.06176985;
      W_o[14,33] := 0.17464209;
      W_o[14,34] := 0.23947489;
      W_o[14,35] := -0.19607270;
      W_o[14,36] := 0.05518134;
      W_o[14,37] := 0.09389904;
      W_o[14,38] := 0.08116579;
      W_o[14,39] := 0.13854055;
      W_o[15,0] := -0.20354150;
      W_o[15,1] := 0.22298840;
      W_o[15,2] := -0.72846305;
      W_o[15,3] := 0.12790513;
      W_o[15,4] := -0.00086900;
      W_o[15,5] := 0.53668076;
      W_o[15,6] := -0.01224643;
      W_o[15,7] := 0.13361789;
      W_o[15,8] := -0.35204136;
      W_o[15,9] := -0.00480295;
      W_o[15,10] := 0.13339433;
      W_o[15,11] := 0.05102095;
      W_o[15,12] := -0.05708028;
      W_o[15,13] := -0.06014942;
      W_o[15,14] := 0.01049514;
      W_o[15,15] := -0.09353844;
      W_o[15,16] := 0.07731096;
      W_o[15,17] := 0.01013883;
      W_o[15,18] := 0.07310723;
      W_o[15,19] := -0.86926681;
      W_o[15,20] := -0.21554285;
      W_o[15,21] := 0.09906635;
      W_o[15,22] := -0.03062510;
      W_o[15,23] := 0.34554279;
      W_o[15,24] := -0.18611832;
      W_o[15,25] := -0.21096791;
      W_o[15,26] := -0.05899647;
      W_o[15,27] := 0.01260784;
      W_o[15,28] := 0.04030582;
      W_o[15,29] := 0.14234707;
      W_o[15,30] := 0.28686827;
      W_o[15,31] := 0.10269888;
      W_o[15,32] := 0.24122585;
      W_o[15,33] := -0.04419544;
      W_o[15,34] := 0.12896782;
      W_o[15,35] := -0.29434389;
      W_o[15,36] := -0.00652304;
      W_o[15,37] := -0.03412445;
      W_o[15,38] := 0.48026237;
      W_o[15,39] := 0.22275838;
      R_i[0,0] := -0.01601154;
      R_i[0,1] := -0.45056638;
      R_i[0,2] := 0.31150612;
      R_i[0,3] := 0.75380063;
      R_i[0,4] := -0.14020784;
      R_i[0,5] := -0.04954997;
      R_i[0,6] := -0.08327835;
      R_i[0,7] := 0.37333494;
      R_i[0,8] := 0.69632649;
      R_i[0,9] := 0.28636262;
      R_i[0,10] := 0.79977125;
      R_i[0,11] := -0.74981761;
      R_i[0,12] := -0.65260571;
      R_i[0,13] := 0.13876246;
      R_i[0,14] := 0.08631746;
      R_i[0,15] := 0.05898035;
      R_i[1,0] := -0.40123200;
      R_i[1,1] := 0.73352093;
      R_i[1,2] := -0.09579885;
      R_i[1,3] := 0.02985846;
      R_i[1,4] := -0.31864849;
      R_i[1,5] := -0.23945375;
      R_i[1,6] := 0.54185194;
      R_i[1,7] := -0.27102774;
      R_i[1,8] := 0.00622073;
      R_i[1,9] := 0.09155256;
      R_i[1,10] := 0.14616042;
      R_i[1,11] := -0.00168930;
      R_i[1,12] := 0.22379795;
      R_i[1,13] := 0.16731951;
      R_i[1,14] := -0.07847317;
      R_i[1,15] := -0.07302959;
      R_i[2,0] := 0.21432666;
      R_i[2,1] := -0.52472848;
      R_i[2,2] := 0.33226553;
      R_i[2,3] := 0.29653755;
      R_i[2,4] := 0.13181669;
      R_i[2,5] := 0.14462742;
      R_i[2,6] := -0.13044202;
      R_i[2,7] := -0.11953641;
      R_i[2,8] := -0.31265071;
      R_i[2,9] := -0.24024297;
      R_i[2,10] := 0.08897854;
      R_i[2,11] := -0.33833930;
      R_i[2,12] := -0.19799015;
      R_i[2,13] := 0.07993159;
      R_i[2,14] := -0.11292934;
      R_i[2,15] := -0.07898453;
      R_i[3,0] := 0.21617912;
      R_i[3,1] := 0.14047004;
      R_i[3,2] := -0.33971104;
      R_i[3,3] := -0.87813431;
      R_i[3,4] := 0.18907729;
      R_i[3,5] := -0.08525109;
      R_i[3,6] := 0.00524858;
      R_i[3,7] := 0.61694282;
      R_i[3,8] := -0.02290213;
      R_i[3,9] := -0.12324939;
      R_i[3,10] := 0.18364368;
      R_i[3,11] := -0.00976140;
      R_i[3,12] := -0.00912099;
      R_i[3,13] := 0.08642489;
      R_i[3,14] := -0.11980756;
      R_i[3,15] := -0.12185419;
      R_i[4,0] := -0.16884419;
      R_i[4,1] := -0.01549527;
      R_i[4,2] := -0.09087992;
      R_i[4,3] := 0.20354238;
      R_i[4,4] := 0.03523245;
      R_i[4,5] := -0.79665762;
      R_i[4,6] := 0.01135984;
      R_i[4,7] := 0.16435672;
      R_i[4,8] := 0.24640194;
      R_i[4,9] := 0.34898201;
      R_i[4,10] := 0.10282461;
      R_i[4,11] := 0.00752686;
      R_i[4,12] := 0.04740289;
      R_i[4,13] := 0.65646058;
      R_i[4,14] := 0.34154060;
      R_i[4,15] := -0.18205808;
      R_i[5,0] := 0.14134005;
      R_i[5,1] := -0.52419472;
      R_i[5,2] := 0.29793712;
      R_i[5,3] := 0.54927635;
      R_i[5,4] := -0.54260975;
      R_i[5,5] := -0.51202631;
      R_i[5,6] := -0.60210627;
      R_i[5,7] := -0.56587559;
      R_i[5,8] := 0.28321642;
      R_i[5,9] := 0.27916816;
      R_i[5,10] := 0.04958420;
      R_i[5,11] := -0.45784742;
      R_i[5,12] := -0.64853847;
      R_i[5,13] := 0.06905902;
      R_i[5,14] := -0.40434125;
      R_i[5,15] := -0.32038039;
      R_i[6,0] := -0.14098248;
      R_i[6,1] := -0.58484751;
      R_i[6,2] := 0.14535309;
      R_i[6,3] := 0.07121052;
      R_i[6,4] := -0.36041209;
      R_i[6,5] := -0.39794296;
      R_i[6,6] := -1.12201309;
      R_i[6,7] := -0.13091828;
      R_i[6,8] := -0.19139199;
      R_i[6,9] := 0.02611434;
      R_i[6,10] := -0.22105527;
      R_i[6,11] := 0.03291342;
      R_i[6,12] := -0.32781577;
      R_i[6,13] := 0.34615195;
      R_i[6,14] := 0.26723450;
      R_i[6,15] := 0.16197382;
      R_i[7,0] := -0.14755228;
      R_i[7,1] := -0.68282712;
      R_i[7,2] := -0.27109590;
      R_i[7,3] := 0.32158145;
      R_i[7,4] := 0.03019373;
      R_i[7,5] := 0.16966243;
      R_i[7,6] := 0.11984173;
      R_i[7,7] := -0.10196535;
      R_i[7,8] := 0.59090692;
      R_i[7,9] := -0.39028153;
      R_i[7,10] := 0.24009976;
      R_i[7,11] := -0.39055178;
      R_i[7,12] := -0.38680884;
      R_i[7,13] := -0.17643671;
      R_i[7,14] := 0.23875171;
      R_i[7,15] := -0.10718834;
      R_i[8,0] := -0.23345003;
      R_i[8,1] := -0.38775986;
      R_i[8,2] := -0.33172470;
      R_i[8,3] := 0.14901052;
      R_i[8,4] := 0.07190004;
      R_i[8,5] := -0.05165868;
      R_i[8,6] := 0.49192744;
      R_i[8,7] := 0.63586611;
      R_i[8,8] := -0.12973778;
      R_i[8,9] := -0.39154807;
      R_i[8,10] := 0.01818666;
      R_i[8,11] := -0.31032625;
      R_i[8,12] := -0.29012892;
      R_i[8,13] := -0.01039465;
      R_i[8,14] := 0.19450903;
      R_i[8,15] := -0.20079081;
      R_i[9,0] := -0.27807117;
      R_i[9,1] := 0.00795646;
      R_i[9,2] := 0.15969256;
      R_i[9,3] := -0.09819215;
      R_i[9,4] := 0.00536336;
      R_i[9,5] := -0.01222592;
      R_i[9,6] := 0.05426886;
      R_i[9,7] := -0.22095288;
      R_i[9,8] := 0.15056732;
      R_i[9,9] := -0.26072544;
      R_i[9,10] := 0.33169287;
      R_i[9,11] := 0.10117077;
      R_i[9,12] := -0.21393171;
      R_i[9,13] := 0.42175838;
      R_i[9,14] := 0.01216281;
      R_i[9,15] := -0.08162050;
      R_i[10,0] := 0.12645799;
      R_i[10,1] := 0.02421534;
      R_i[10,2] := -0.24892592;
      R_i[10,3] := 0.09164374;
      R_i[10,4] := -0.42948586;
      R_i[10,5] := -0.05434940;
      R_i[10,6] := 0.56467527;
      R_i[10,7] := 0.33178699;
      R_i[10,8] := 0.26021555;
      R_i[10,9] := -0.39298084;
      R_i[10,10] := -0.39579603;
      R_i[10,11] := -0.00741246;
      R_i[10,12] := -0.33583519;
      R_i[10,13] := -0.01858520;
      R_i[10,14] := 0.44103009;
      R_i[10,15] := -0.09651927;
      R_i[11,0] := 0.09693456;
      R_i[11,1] := -0.35125014;
      R_i[11,2] := -0.02015482;
      R_i[11,3] := 0.35720971;
      R_i[11,4] := -0.11965420;
      R_i[11,5] := 0.14459991;
      R_i[11,6] := -0.19067928;
      R_i[11,7] := 0.08080416;
      R_i[11,8] := 0.17797850;
      R_i[11,9] := -0.14250341;
      R_i[11,10] := -0.38627943;
      R_i[11,11] := 0.49561632;
      R_i[11,12] := -0.17909285;
      R_i[11,13] := 0.20836362;
      R_i[11,14] := 0.40069145;
      R_i[11,15] := 0.38960215;
      R_i[12,0] := 0.34008914;
      R_i[12,1] := -0.17271595;
      R_i[12,2] := -0.30769649;
      R_i[12,3] := -0.28230789;
      R_i[12,4] := 0.05254490;
      R_i[12,5] := 0.07448359;
      R_i[12,6] := -0.00981909;
      R_i[12,7] := 0.10081543;
      R_i[12,8] := 0.30097830;
      R_i[12,9] := 0.29120073;
      R_i[12,10] := 0.12718941;
      R_i[12,11] := -0.06783659;
      R_i[12,12] := 0.44559616;
      R_i[12,13] := -0.32429484;
      R_i[12,14] := -0.18343198;
      R_i[12,15] := -0.10893025;
      R_i[13,0] := -0.28948510;
      R_i[13,1] := -0.16649665;
      R_i[13,2] := 0.04430598;
      R_i[13,3] := 0.11078570;
      R_i[13,4] := -0.56880260;
      R_i[13,5] := -0.07979194;
      R_i[13,6] := 0.15275165;
      R_i[13,7] := 0.12733753;
      R_i[13,8] := 0.36211529;
      R_i[13,9] := 0.30433327;
      R_i[13,10] := -0.17985806;
      R_i[13,11] := -0.23772895;
      R_i[13,12] := 0.12355826;
      R_i[13,13] := 0.50354385;
      R_i[13,14] := 0.10862395;
      R_i[13,15] := -0.02580172;
      R_i[14,0] := 0.04543614;
      R_i[14,1] := -0.40430877;
      R_i[14,2] := 0.12097509;
      R_i[14,3] := 0.48837635;
      R_i[14,4] := 0.00980398;
      R_i[14,5] := 0.03799421;
      R_i[14,6] := 0.32785147;
      R_i[14,7] := 0.06604390;
      R_i[14,8] := 0.17208503;
      R_i[14,9] := -0.37074247;
      R_i[14,10] := -0.13859139;
      R_i[14,11] := 0.27189708;
      R_i[14,12] := -0.13288878;
      R_i[14,13] := 0.27018747;
      R_i[14,14] := 1.38667846;
      R_i[14,15] := 0.05095792;
      R_i[15,0] := 0.12141960;
      R_i[15,1] := -0.03100028;
      R_i[15,2] := 0.26846337;
      R_i[15,3] := 0.21032426;
      R_i[15,4] := -0.11904223;
      R_i[15,5] := 0.09452529;
      R_i[15,6] := 0.30823541;
      R_i[15,7] := -0.00003856;
      R_i[15,8] := 0.27272546;
      R_i[15,9] := 0.05441154;
      R_i[15,10] := -0.12308154;
      R_i[15,11] := -0.47818425;
      R_i[15,12] := -0.21431655;
      R_i[15,13] := -0.24715155;
      R_i[15,14] := 0.20871881;
      R_i[15,15] := 0.02325043;
      R_f[0,0] := -0.03493118;
      R_f[0,1] := -0.37833330;
      R_f[0,2] := 0.03728793;
      R_f[0,3] := 0.14278547;
      R_f[0,4] := -0.12003965;
      R_f[0,5] := -0.06856227;
      R_f[0,6] := 0.07930882;
      R_f[0,7] := 0.27766067;
      R_f[0,8] := 0.07494716;
      R_f[0,9] := 0.14615805;
      R_f[0,10] := -0.07652009;
      R_f[0,11] := -0.09052465;
      R_f[0,12] := -0.11576622;
      R_f[0,13] := 0.04987612;
      R_f[0,14] := 0.06529343;
      R_f[0,15] := 0.00263772;
      R_f[1,0] := -0.43777743;
      R_f[1,1] := 0.72514027;
      R_f[1,2] := -0.38771391;
      R_f[1,3] := -0.01443690;
      R_f[1,4] := -0.00149874;
      R_f[1,5] := -0.34476724;
      R_f[1,6] := 0.29173759;
      R_f[1,7] := 0.09541123;
      R_f[1,8] := 0.34579757;
      R_f[1,9] := 0.62985712;
      R_f[1,10] := 0.05302448;
      R_f[1,11] := 0.20725778;
      R_f[1,12] := -0.04234733;
      R_f[1,13] := 0.33368251;
      R_f[1,14] := 0.13071071;
      R_f[1,15] := 0.12571791;
      R_f[2,0] := 0.33107671;
      R_f[2,1] := -0.38107035;
      R_f[2,2] := 0.11539750;
      R_f[2,3] := 0.34765753;
      R_f[2,4] := -0.24806751;
      R_f[2,5] := 0.12396693;
      R_f[2,6] := -0.00015690;
      R_f[2,7] := -0.03111286;
      R_f[2,8] := -0.40619534;
      R_f[2,9] := -0.10276131;
      R_f[2,10] := -0.01848604;
      R_f[2,11] := -0.38150114;
      R_f[2,12] := 0.07561549;
      R_f[2,13] := -0.32942322;
      R_f[2,14] := -0.04146929;
      R_f[2,15] := 0.10218077;
      R_f[3,0] := -0.95647854;
      R_f[3,1] := 0.32638514;
      R_f[3,2] := -0.18242189;
      R_f[3,3] := -0.29949248;
      R_f[3,4] := 0.17140226;
      R_f[3,5] := -0.20921187;
      R_f[3,6] := -0.10329774;
      R_f[3,7] := -0.15821460;
      R_f[3,8] := 0.15070482;
      R_f[3,9] := 0.33798599;
      R_f[3,10] := -0.27949187;
      R_f[3,11] := 0.08474356;
      R_f[3,12] := 0.24811046;
      R_f[3,13] := 0.09939278;
      R_f[3,14] := -0.24101312;
      R_f[3,15] := -0.19353758;
      R_f[4,0] := -0.23498796;
      R_f[4,1] := -0.40744987;
      R_f[4,2] := 0.26351565;
      R_f[4,3] := -0.26684532;
      R_f[4,4] := -0.09082807;
      R_f[4,5] := -0.08405253;
      R_f[4,6] := 0.08696185;
      R_f[4,7] := 0.11129832;
      R_f[4,8] := 0.16387634;
      R_f[4,9] := -0.11868069;
      R_f[4,10] := 0.32621741;
      R_f[4,11] := -0.14263494;
      R_f[4,12] := 0.13083991;
      R_f[4,13] := 0.17955558;
      R_f[4,14] := 0.16594826;
      R_f[4,15] := 0.12359417;
      R_f[5,0] := 0.35480824;
      R_f[5,1] := -0.12709811;
      R_f[5,2] := 0.24268471;
      R_f[5,3] := 0.08011950;
      R_f[5,4] := 0.21156235;
      R_f[5,5] := 0.27579746;
      R_f[5,6] := 0.20017114;
      R_f[5,7] := 0.01883883;
      R_f[5,8] := -0.39427981;
      R_f[5,9] := -0.35867786;
      R_f[5,10] := 0.06389395;
      R_f[5,11] := -0.11106856;
      R_f[5,12] := 0.11757033;
      R_f[5,13] := -0.01875320;
      R_f[5,14] := 0.01303833;
      R_f[5,15] := -0.06690010;
      R_f[6,0] := -0.50047231;
      R_f[6,1] := -0.07684148;
      R_f[6,2] := 0.19817993;
      R_f[6,3] := 0.05971020;
      R_f[6,4] := -0.04680483;
      R_f[6,5] := 0.31770298;
      R_f[6,6] := 0.12533610;
      R_f[6,7] := 0.13815877;
      R_f[6,8] := 0.02148284;
      R_f[6,9] := -0.06106690;
      R_f[6,10] := 0.13362114;
      R_f[6,11] := 0.21636069;
      R_f[6,12] := -0.09828766;
      R_f[6,13] := 0.21644033;
      R_f[6,14] := 0.20338993;
      R_f[6,15] := 0.14178181;
      R_f[7,0] := 0.26125121;
      R_f[7,1] := -0.03714739;
      R_f[7,2] := 0.08117681;
      R_f[7,3] := 0.20744996;
      R_f[7,4] := -0.32044601;
      R_f[7,5] := 0.41264480;
      R_f[7,6] := 0.61615700;
      R_f[7,7] := -0.17647557;
      R_f[7,8] := -0.15667132;
      R_f[7,9] := -0.02732511;
      R_f[7,10] := -0.49891508;
      R_f[7,11] := 0.00061774;
      R_f[7,12] := -0.02982556;
      R_f[7,13] := 0.03914607;
      R_f[7,14] := 0.20352171;
      R_f[7,15] := 0.01521025;
      R_f[8,0] := -0.00262567;
      R_f[8,1] := -0.19572628;
      R_f[8,2] := -0.01333520;
      R_f[8,3] := 0.13264976;
      R_f[8,4] := -0.06475109;
      R_f[8,5] := 0.27500546;
      R_f[8,6] := 0.29358950;
      R_f[8,7] := 0.10781989;
      R_f[8,8] := -0.55418187;
      R_f[8,9] := -0.03762578;
      R_f[8,10] := -0.25193849;
      R_f[8,11] := 0.27721903;
      R_f[8,12] := -0.15396175;
      R_f[8,13] := -0.02145483;
      R_f[8,14] := 0.24167821;
      R_f[8,15] := 0.06824671;
      R_f[9,0] := 0.25040591;
      R_f[9,1] := -0.33838606;
      R_f[9,2] := 0.06741230;
      R_f[9,3] := 0.20970462;
      R_f[9,4] := -0.08986910;
      R_f[9,5] := -0.20913272;
      R_f[9,6] := 0.31628108;
      R_f[9,7] := 0.26534095;
      R_f[9,8] := 0.02326944;
      R_f[9,9] := -0.80536783;
      R_f[9,10] := -0.24160722;
      R_f[9,11] := -0.03336972;
      R_f[9,12] := -0.36345491;
      R_f[9,13] := 0.01661946;
      R_f[9,14] := -0.11790104;
      R_f[9,15] := 0.14004685;
      R_f[10,0] := 0.20252159;
      R_f[10,1] := -0.33094549;
      R_f[10,2] := 0.28349048;
      R_f[10,3] := 0.20983174;
      R_f[10,4] := -0.39166585;
      R_f[10,5] := 0.14894433;
      R_f[10,6] := 0.05038162;
      R_f[10,7] := 0.14217970;
      R_f[10,8] := -0.24751066;
      R_f[10,9] := 0.04759743;
      R_f[10,10] := -0.16426384;
      R_f[10,11] := -0.16217081;
      R_f[10,12] := -0.12350682;
      R_f[10,13] := 0.08995254;
      R_f[10,14] := -0.01327613;
      R_f[10,15] := 0.22854908;
      R_f[11,0] := 0.16012208;
      R_f[11,1] := 0.26288185;
      R_f[11,2] := 0.21906035;
      R_f[11,3] := -0.04701964;
      R_f[11,4] := -0.13884930;
      R_f[11,5] := 0.08709867;
      R_f[11,6] := -0.07009537;
      R_f[11,7] := -0.16951092;
      R_f[11,8] := 0.02868164;
      R_f[11,9] := -0.01121150;
      R_f[11,10] := 0.07267684;
      R_f[11,11] := -0.19895513;
      R_f[11,12] := 0.36136580;
      R_f[11,13] := -0.05935945;
      R_f[11,14] := 0.08223550;
      R_f[11,15] := 0.37379497;
      R_f[12,0] := -0.25996360;
      R_f[12,1] := -0.48404145;
      R_f[12,2] := -0.32950810;
      R_f[12,3] := 0.11100189;
      R_f[12,4] := -0.26770976;
      R_f[12,5] := -0.17353055;
      R_f[12,6] := 0.16970958;
      R_f[12,7] := -0.34763816;
      R_f[12,8] := 0.51724803;
      R_f[12,9] := -0.22855559;
      R_f[12,10] := 0.86062002;
      R_f[12,11] := 0.06095523;
      R_f[12,12] := -0.12677126;
      R_f[12,13] := 0.23355845;
      R_f[12,14] := 0.24020465;
      R_f[12,15] := -0.22797880;
      R_f[13,0] := 0.02567713;
      R_f[13,1] := -0.31515360;
      R_f[13,2] := -0.12621829;
      R_f[13,3] := 0.18368529;
      R_f[13,4] := -0.03905401;
      R_f[13,5] := 0.71356320;
      R_f[13,6] := 0.08130559;
      R_f[13,7] := 0.01576971;
      R_f[13,8] := -0.20504172;
      R_f[13,9] := 0.07079811;
      R_f[13,10] := -0.10902814;
      R_f[13,11] := 0.15747260;
      R_f[13,12] := -0.34046116;
      R_f[13,13] := 0.10420194;
      R_f[13,14] := -0.05406023;
      R_f[13,15] := 0.23026128;
      R_f[14,0] := 0.05553682;
      R_f[14,1] := 0.03039004;
      R_f[14,2] := -0.39775774;
      R_f[14,3] := 0.17736661;
      R_f[14,4] := -0.14014874;
      R_f[14,5] := 0.18136151;
      R_f[14,6] := 0.08784663;
      R_f[14,7] := -0.00406716;
      R_f[14,8] := 0.29372466;
      R_f[14,9] := -0.21857265;
      R_f[14,10] := 0.32868984;
      R_f[14,11] := 0.52028972;
      R_f[14,12] := 0.27974731;
      R_f[14,13] := -0.10954703;
      R_f[14,14] := 1.17473233;
      R_f[14,15] := 0.29271725;
      R_f[15,0] := 0.35421464;
      R_f[15,1] := -0.62420565;
      R_f[15,2] := 0.22943251;
      R_f[15,3] := 0.29831216;
      R_f[15,4] := -0.20180914;
      R_f[15,5] := 0.39882076;
      R_f[15,6] := 0.27627981;
      R_f[15,7] := 0.38468793;
      R_f[15,8] := 0.04349254;
      R_f[15,9] := -0.10810658;
      R_f[15,10] := -0.37345368;
      R_f[15,11] := -0.10984580;
      R_f[15,12] := 0.33647370;
      R_f[15,13] := 0.34551468;
      R_f[15,14] := 0.02944022;
      R_f[15,15] := 0.02307001;
      R_g[0,0] := -1.25112379;
      R_g[0,1] := -0.21883342;
      R_g[0,2] := 0.11012935;
      R_g[0,3] := 0.25012675;
      R_g[0,4] := -0.10405856;
      R_g[0,5] := 0.13891214;
      R_g[0,6] := 0.10241263;
      R_g[0,7] := 0.22247586;
      R_g[0,8] := 0.06886309;
      R_g[0,9] := -0.05504098;
      R_g[0,10] := 0.13162677;
      R_g[0,11] := -0.09226879;
      R_g[0,12] := 0.03665201;
      R_g[0,13] := 0.01448225;
      R_g[0,14] := 0.08514914;
      R_g[0,15] := 0.10349822;
      R_g[1,0] := -0.01289242;
      R_g[1,1] := -0.76937956;
      R_g[1,2] := -0.00765862;
      R_g[1,3] := -0.02182954;
      R_g[1,4] := -0.00624790;
      R_g[1,5] := -0.09856889;
      R_g[1,6] := -0.00179921;
      R_g[1,7] := -0.15975930;
      R_g[1,8] := 0.14410421;
      R_g[1,9] := -0.13659404;
      R_g[1,10] := -0.10461834;
      R_g[1,11] := 0.17878979;
      R_g[1,12] := 0.13712661;
      R_g[1,13] := 0.10399450;
      R_g[1,14] := 0.20643574;
      R_g[1,15] := 0.05955669;
      R_g[2,0] := -0.00450423;
      R_g[2,1] := 0.27837455;
      R_g[2,2] := -1.65240133;
      R_g[2,3] := -0.08348246;
      R_g[2,4] := 0.00295603;
      R_g[2,5] := -0.12203792;
      R_g[2,6] := -0.01780931;
      R_g[2,7] := 0.08614038;
      R_g[2,8] := -0.05562058;
      R_g[2,9] := 0.10056782;
      R_g[2,10] := 0.03247114;
      R_g[2,11] := -0.11223084;
      R_g[2,12] := -0.10098543;
      R_g[2,13] := 0.01667355;
      R_g[2,14] := -0.26046327;
      R_g[2,15] := -0.26248303;
      R_g[3,0] := -0.03127015;
      R_g[3,1] := 0.23647039;
      R_g[3,2] := -0.25464910;
      R_g[3,3] := -0.99465227;
      R_g[3,4] := -0.00474326;
      R_g[3,5] := 0.02257820;
      R_g[3,6] := -0.12011071;
      R_g[3,7] := -0.36244613;
      R_g[3,8] := 0.16971782;
      R_g[3,9] := 0.18556982;
      R_g[3,10] := 0.12659717;
      R_g[3,11] := -0.07901487;
      R_g[3,12] := -0.08990744;
      R_g[3,13] := 0.14218350;
      R_g[3,14] := -0.14387904;
      R_g[3,15] := -0.29380691;
      R_g[4,0] := 0.07746305;
      R_g[4,1] := 0.05525218;
      R_g[4,2] := 0.18610036;
      R_g[4,3] := 0.11015689;
      R_g[4,4] := -1.79593194;
      R_g[4,5] := -0.03749003;
      R_g[4,6] := 0.01035422;
      R_g[4,7] := 0.10059743;
      R_g[4,8] := 0.23833929;
      R_g[4,9] := -0.04896057;
      R_g[4,10] := -0.10350814;
      R_g[4,11] := 0.05637380;
      R_g[4,12] := -0.25450024;
      R_g[4,13] := -0.08886177;
